// CFC twin of T_SafeEStop_Tests: the same tests drawn as CFC diagrams, the way a TwinSAFE project is authored.
    FUNCTION_BLOCK T_SafeEStop_Tests_CFC EXTENDS T_SafeCfcTestSuite
    VAR
    // Test_OutputsOffWhenStopped
    group_1 : T_SafeGroup;
    fb_1 : T_SafeEStop(group := group_1);
    // Test_StartupRequiresRestartSequence
    group_2 : T_SafeGroup;
    fb_2 : T_SafeEStop(group := group_2);
    // Test_EStopRequestSwitchesOutputsOffAndBlocksRestart
    group_3 : T_SafeGroup;
    fb_3 : T_SafeEStop(group := group_3);
    // Test_MakeContactInputRequestsSafeStateOnOne
    group_4 : T_SafeGroup;
    fb_4 : T_SafeEStop(group := group_4) := (Parameters := (EStopIn1MakeContact := TRUE));
    // Test_EdmErrorAtRestartAndAcknowledge
    group_5 : T_SafeGroup;
    fb_5 : T_SafeEStop(group := group_5);
    // Test_RestartHeldBeforeEStopGivesEdmError
    group_6 : T_SafeGroup;
    fb_6 : T_SafeEStop(group := group_6);
    // Test_DelayedOutput
    group_7 : T_SafeGroup;
    fb_7 : T_SafeEStop(group := group_7) := (Parameters := (DelayTime := T#150MS));
    tR1_7 : TON;
    tR2_7 : TON;
    tPress_7 : TON;
    t1_7 : TON;
    trigPress_7 : R_TRIG;
    trig1_7 : R_TRIG;
    // Test_DiscrepancyErrorNeedsSafeInputsBeforeAck
    group_8 : T_SafeGroup;
    fb_8 : T_SafeEStop(group := group_8) := (Parameters := (DiscrepancyTime1 := T#100MS));
    tR1_8 : TON;
    tR2_8 : TON;
    tPress_8 : TON;
    t1_8 : TON;
    trig1_8 : R_TRIG;
END_VAR

Test_OutputsOffWhenStopped();
Test_StartupRequiresRestartSequence();
Test_EStopRequestSwitchesOutputsOffAndBlocksRestart();
Test_MakeContactInputRequestsSafeStateOnOne();
Test_EdmErrorAtRestartAndAcknowledge();
Test_RestartHeldBeforeEStopGivesEdmError();
Test_DelayedOutput();
Test_DiscrepancyErrorNeedsSafeInputsBeforeAck();

METHOD PRIVATE Test_OutputsOffWhenStopped
// note: this text did not pass the execution check against the stored diagram
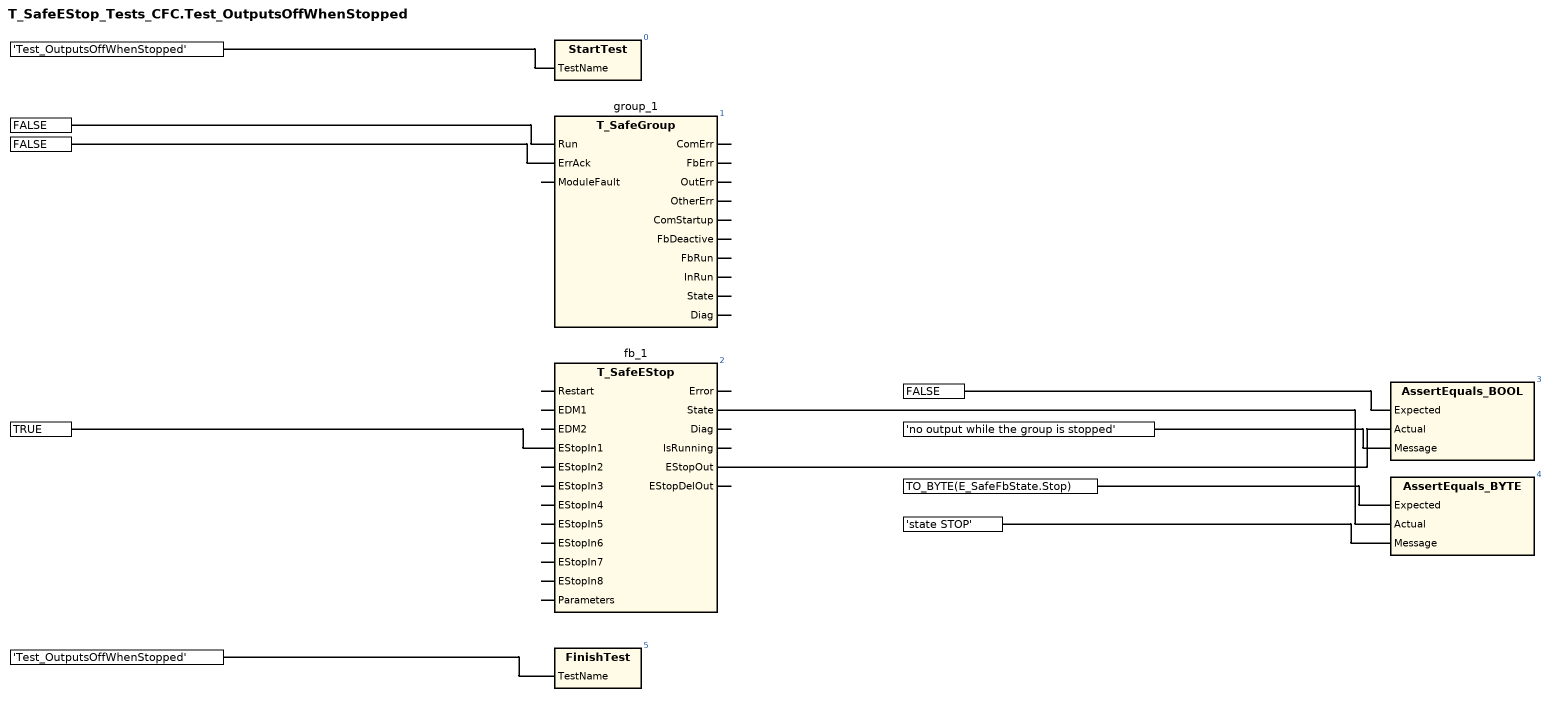
StartTest(TestName := 'Test_OutputsOffWhenStopped');
group_1(Run := FALSE, ErrAck := FALSE); // T_SafeGroup
fb_1(EStopIn1 := TRUE); // T_SafeEStop
AssertEquals_BOOL(Expected := FALSE, Actual := fb_1.EStopOut, Message := 'no output while the group is stopped');
AssertEquals_BYTE(Expected := TO_BYTE(E_SafeFbState.Stop), Actual := fb_1.State, Message := 'state STOP');
FinishTest(TestName := 'Test_OutputsOffWhenStopped');
END_METHOD

METHOD PRIVATE Test_StartupRequiresRestartSequence
// note: this text did not pass the execution check against the stored diagram
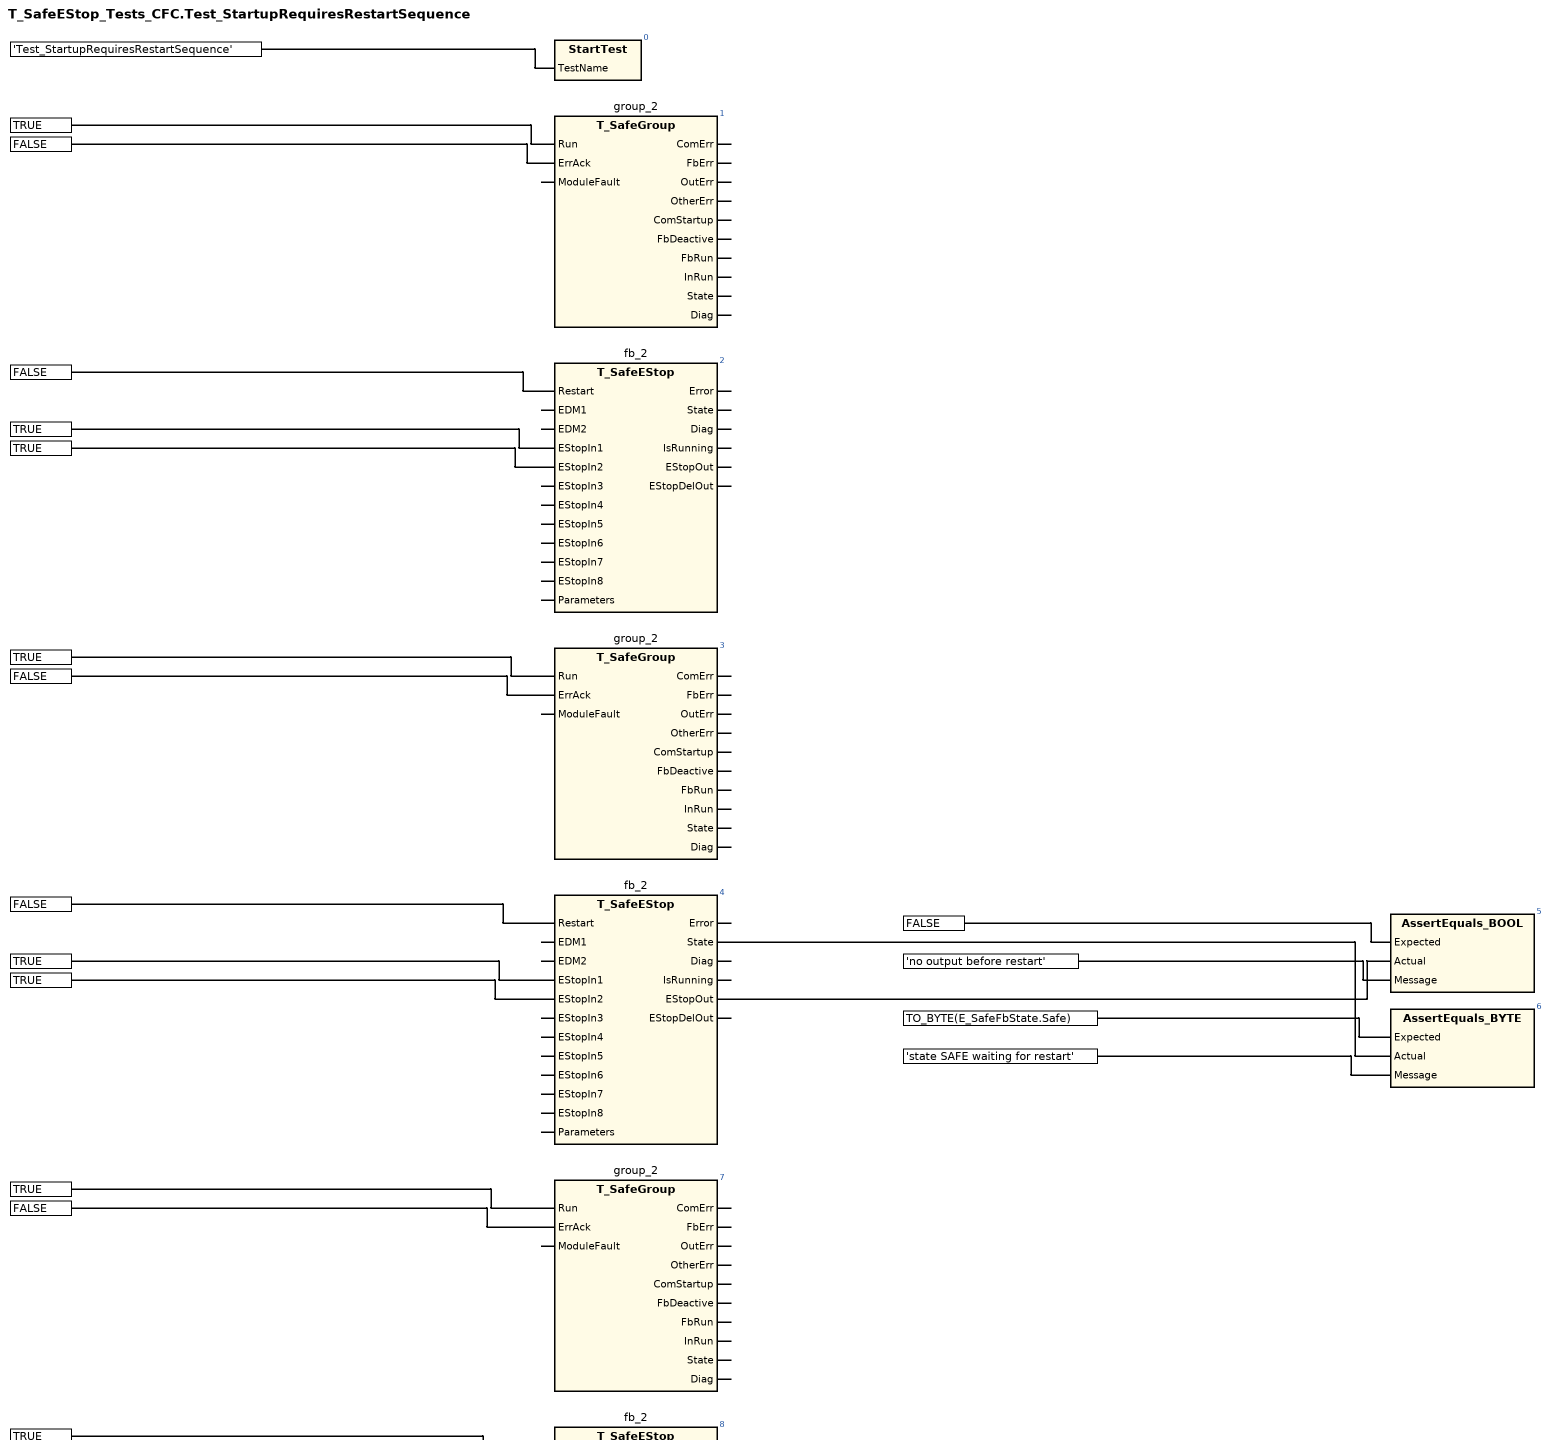
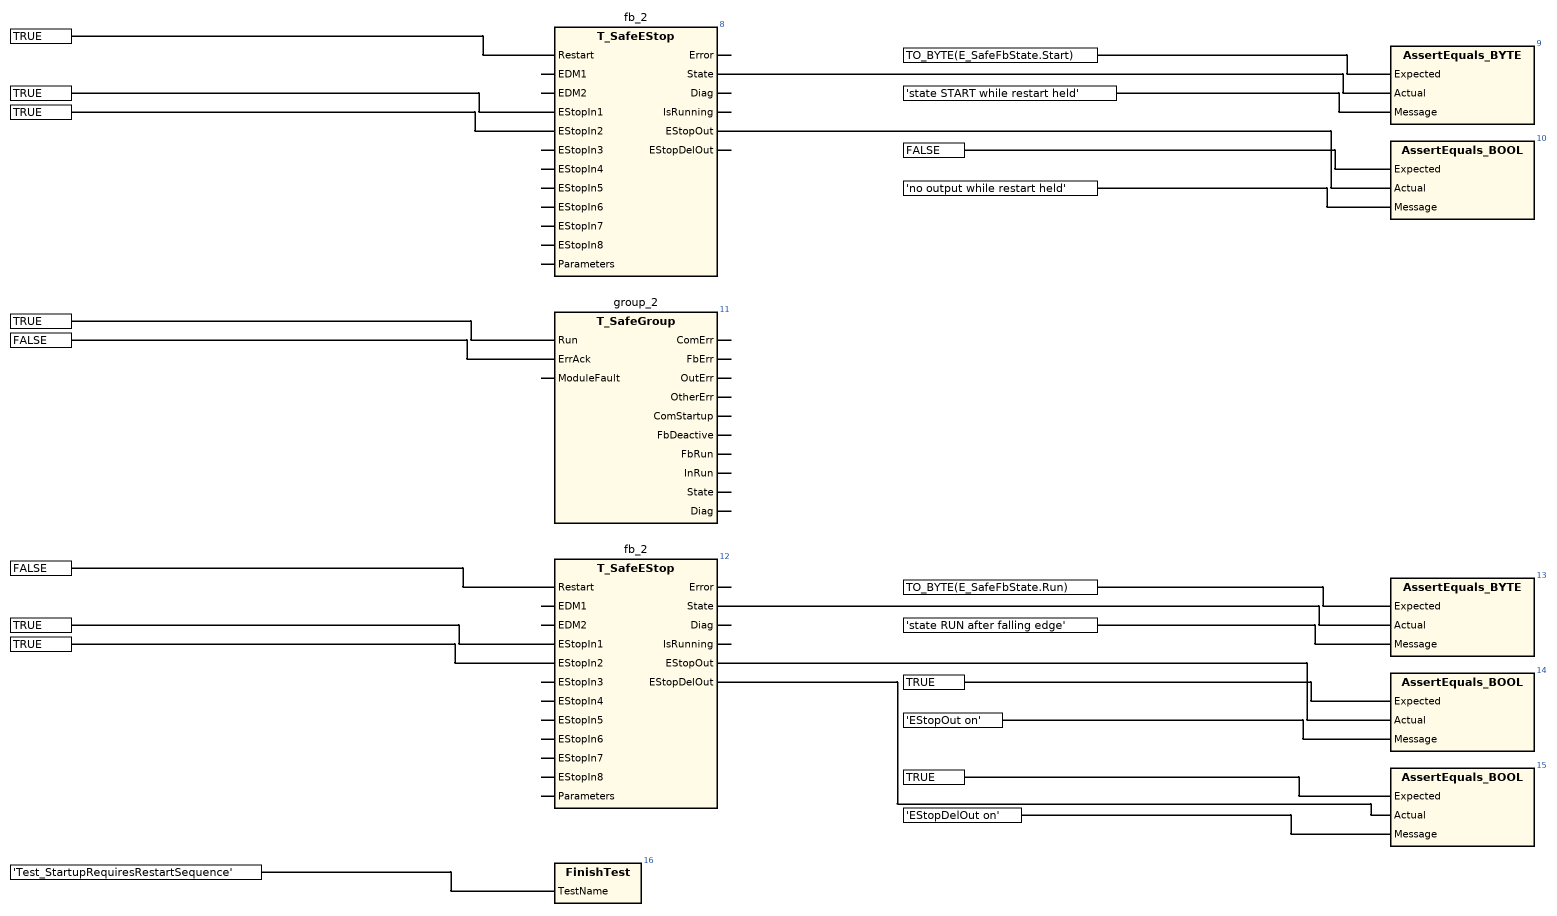
StartTest(TestName := 'Test_StartupRequiresRestartSequence');
group_2(Run := TRUE, ErrAck := FALSE); // T_SafeGroup
fb_2(Restart := FALSE, EStopIn1 := TRUE, EStopIn2 := TRUE); // T_SafeEStop
group_2(Run := TRUE, ErrAck := FALSE); // T_SafeGroup
fb_2(Restart := FALSE, EStopIn1 := TRUE, EStopIn2 := TRUE); // T_SafeEStop
AssertEquals_BOOL(Expected := FALSE, Actual := fb_2.EStopOut, Message := 'no output before restart');
AssertEquals_BYTE(Expected := TO_BYTE(E_SafeFbState.Safe), Actual := fb_2.State, Message := 'state SAFE waiting for restart');
group_2(Run := TRUE, ErrAck := FALSE); // T_SafeGroup
fb_2(Restart := TRUE, EStopIn1 := TRUE, EStopIn2 := TRUE); // T_SafeEStop
AssertEquals_BYTE(Expected := TO_BYTE(E_SafeFbState.Start), Actual := fb_2.State, Message := 'state START while restart held');
AssertEquals_BOOL(Expected := FALSE, Actual := fb_2.EStopOut, Message := 'no output while restart held');
group_2(Run := TRUE, ErrAck := FALSE); // T_SafeGroup
fb_2(Restart := FALSE, EStopIn1 := TRUE, EStopIn2 := TRUE); // T_SafeEStop
AssertEquals_BYTE(Expected := TO_BYTE(E_SafeFbState.Run), Actual := fb_2.State, Message := 'state RUN after falling edge');
AssertEquals_BOOL(Expected := TRUE, Actual := fb_2.EStopOut, Message := 'EStopOut on');
AssertEquals_BOOL(Expected := TRUE, Actual := fb_2.EStopDelOut, Message := 'EStopDelOut on');
FinishTest(TestName := 'Test_StartupRequiresRestartSequence');
END_METHOD

METHOD PRIVATE Test_EStopRequestSwitchesOutputsOffAndBlocksRestart
// note: this text did not pass the execution check against the stored diagram
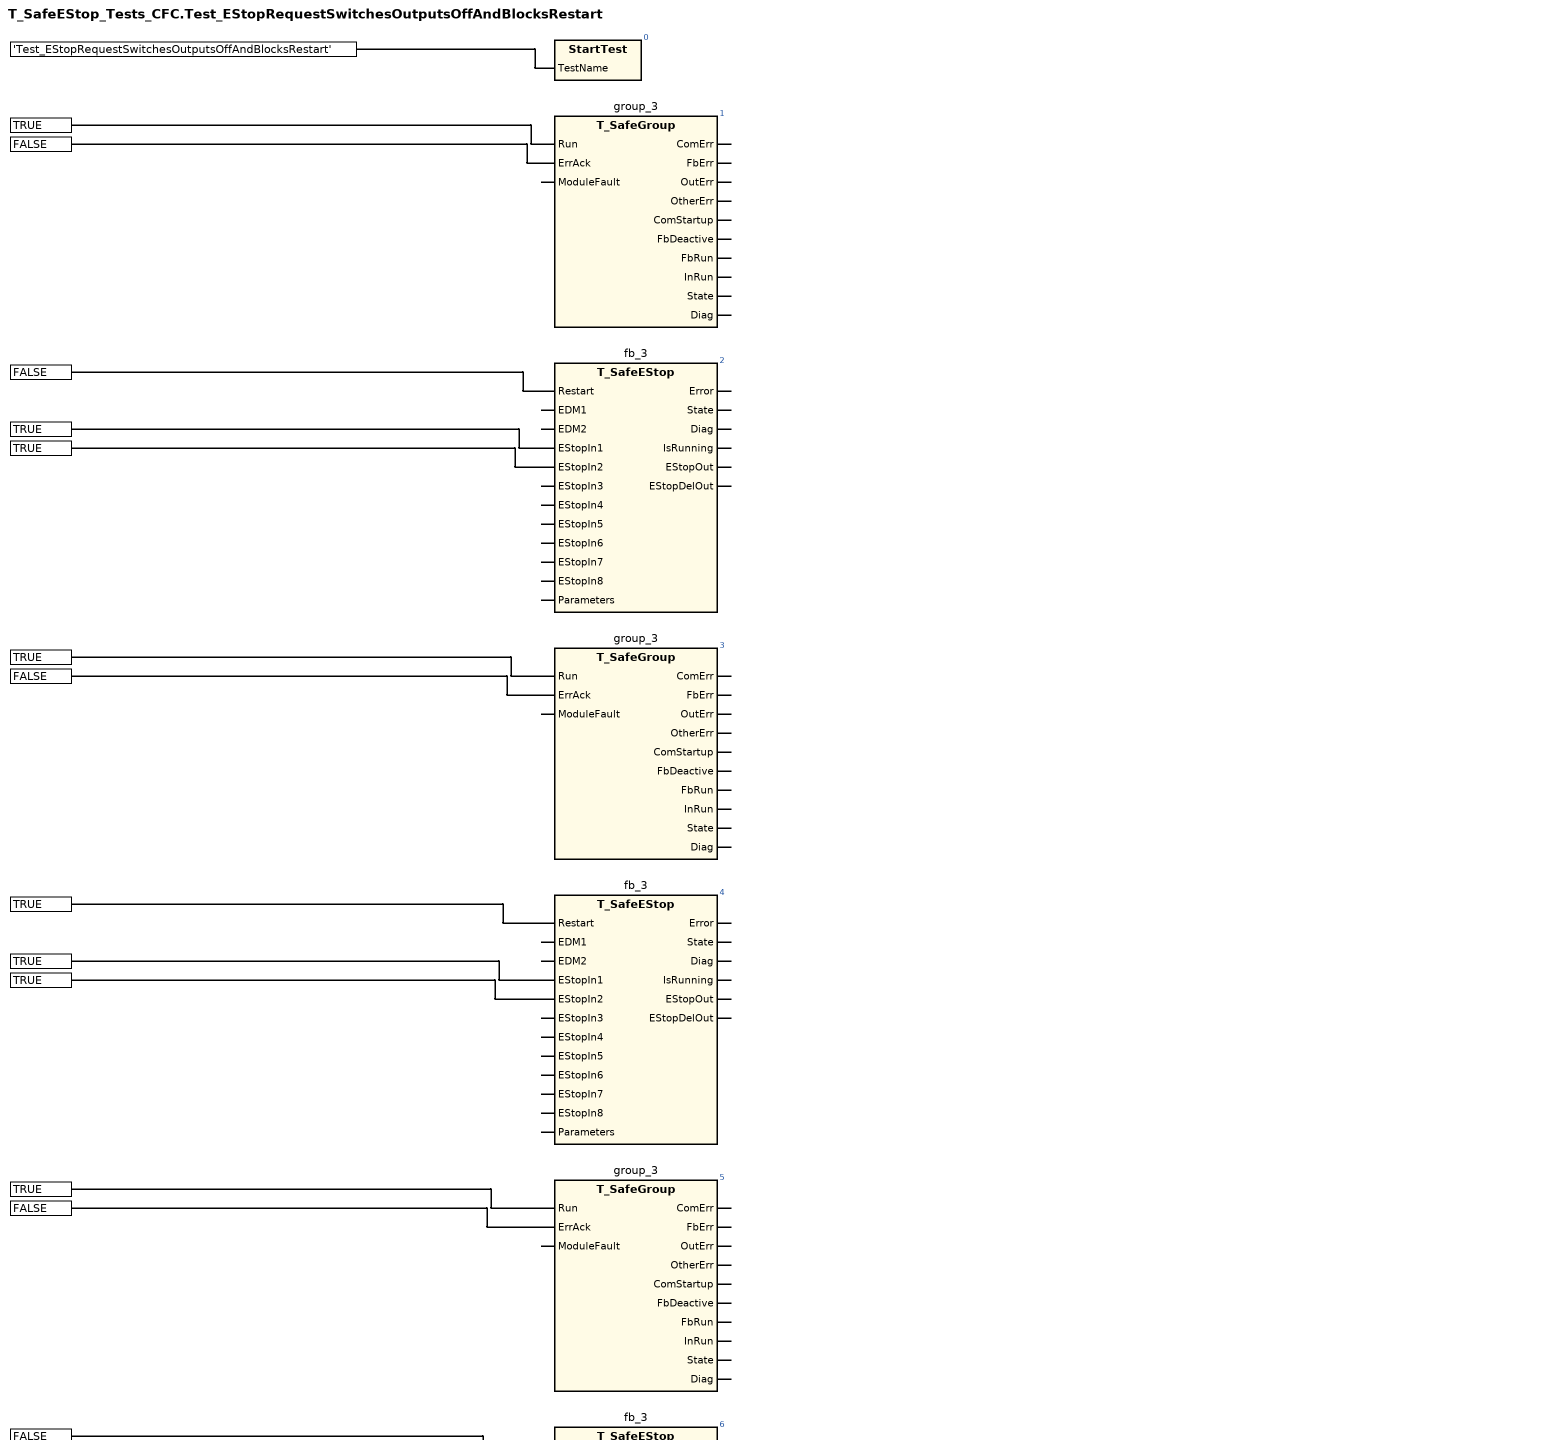
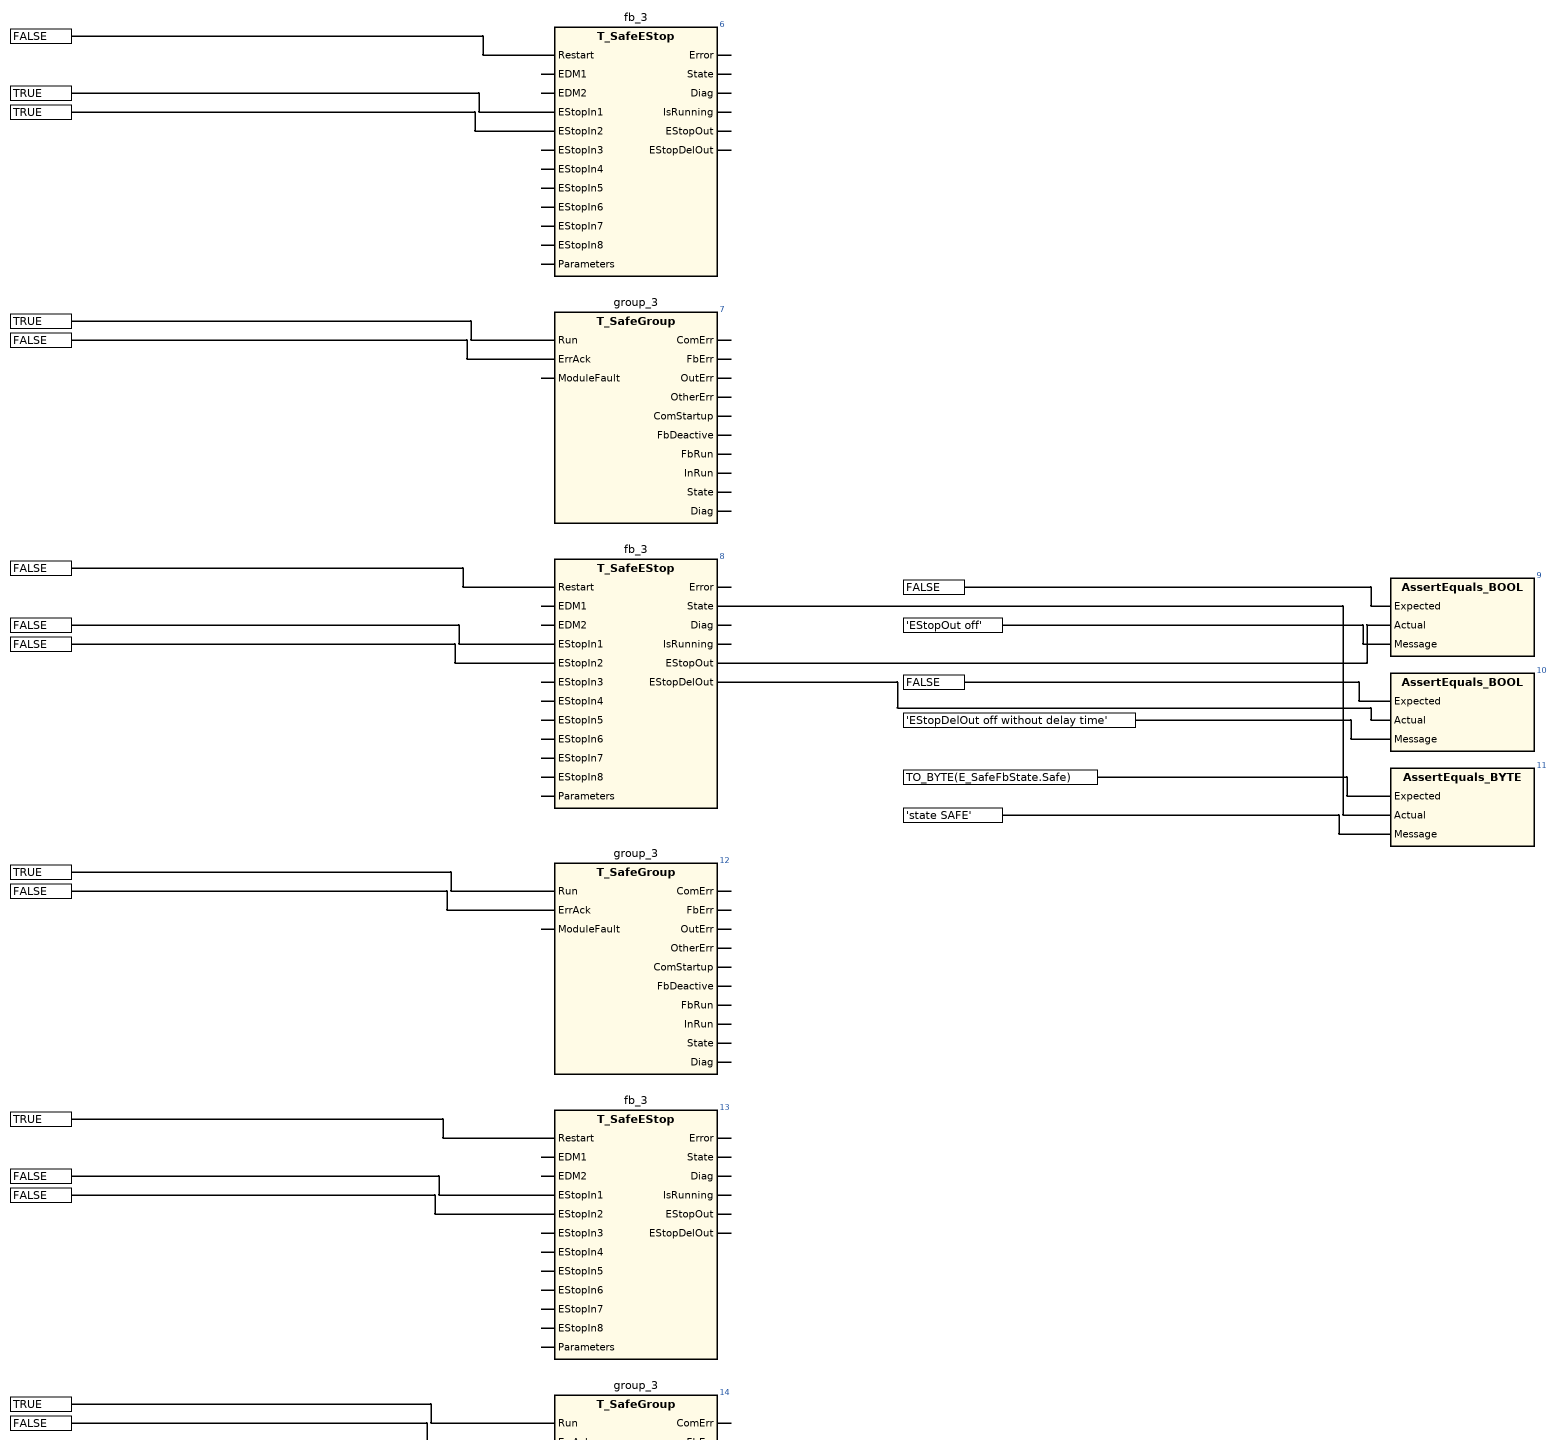
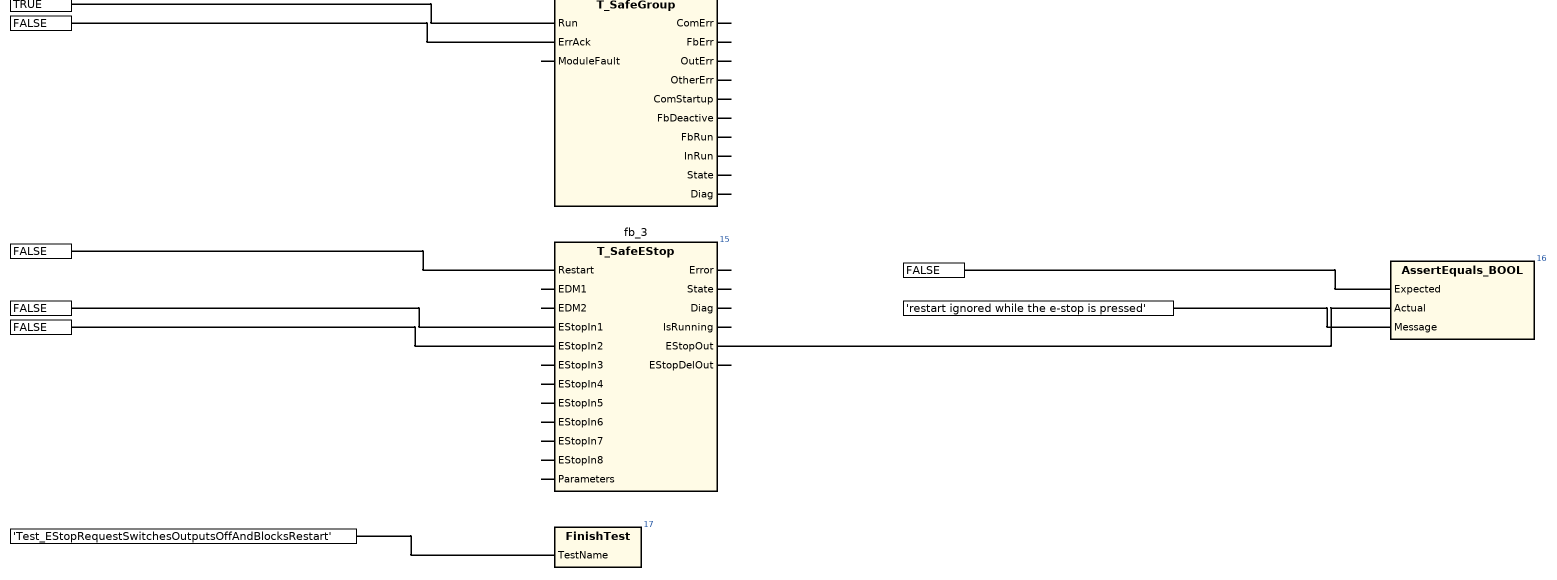
StartTest(TestName := 'Test_EStopRequestSwitchesOutputsOffAndBlocksRestart');
group_3(Run := TRUE, ErrAck := FALSE); // T_SafeGroup
fb_3(Restart := FALSE, EStopIn1 := TRUE, EStopIn2 := TRUE); // T_SafeEStop
group_3(Run := TRUE, ErrAck := FALSE); // T_SafeGroup
fb_3(Restart := TRUE, EStopIn1 := TRUE, EStopIn2 := TRUE); // T_SafeEStop
group_3(Run := TRUE, ErrAck := FALSE); // T_SafeGroup
fb_3(Restart := FALSE, EStopIn1 := TRUE, EStopIn2 := TRUE); // T_SafeEStop
group_3(Run := TRUE, ErrAck := FALSE); // T_SafeGroup
fb_3(Restart := FALSE, EStopIn1 := FALSE, EStopIn2 := FALSE); // T_SafeEStop
AssertEquals_BOOL(Expected := FALSE, Actual := fb_3.EStopOut, Message := 'EStopOut off');
AssertEquals_BOOL(Expected := FALSE, Actual := fb_3.EStopDelOut, Message := 'EStopDelOut off without delay time');
AssertEquals_BYTE(Expected := TO_BYTE(E_SafeFbState.Safe), Actual := fb_3.State, Message := 'state SAFE');
group_3(Run := TRUE, ErrAck := FALSE); // T_SafeGroup
fb_3(Restart := TRUE, EStopIn1 := FALSE, EStopIn2 := FALSE); // T_SafeEStop
group_3(Run := TRUE, ErrAck := FALSE); // T_SafeGroup
fb_3(Restart := FALSE, EStopIn1 := FALSE, EStopIn2 := FALSE); // T_SafeEStop
AssertEquals_BOOL(Expected := FALSE, Actual := fb_3.EStopOut, Message := 'restart ignored while the e-stop is pressed');
FinishTest(TestName := 'Test_EStopRequestSwitchesOutputsOffAndBlocksRestart');
END_METHOD

METHOD PRIVATE Test_MakeContactInputRequestsSafeStateOnOne
// note: this text did not pass the execution check against the stored diagram
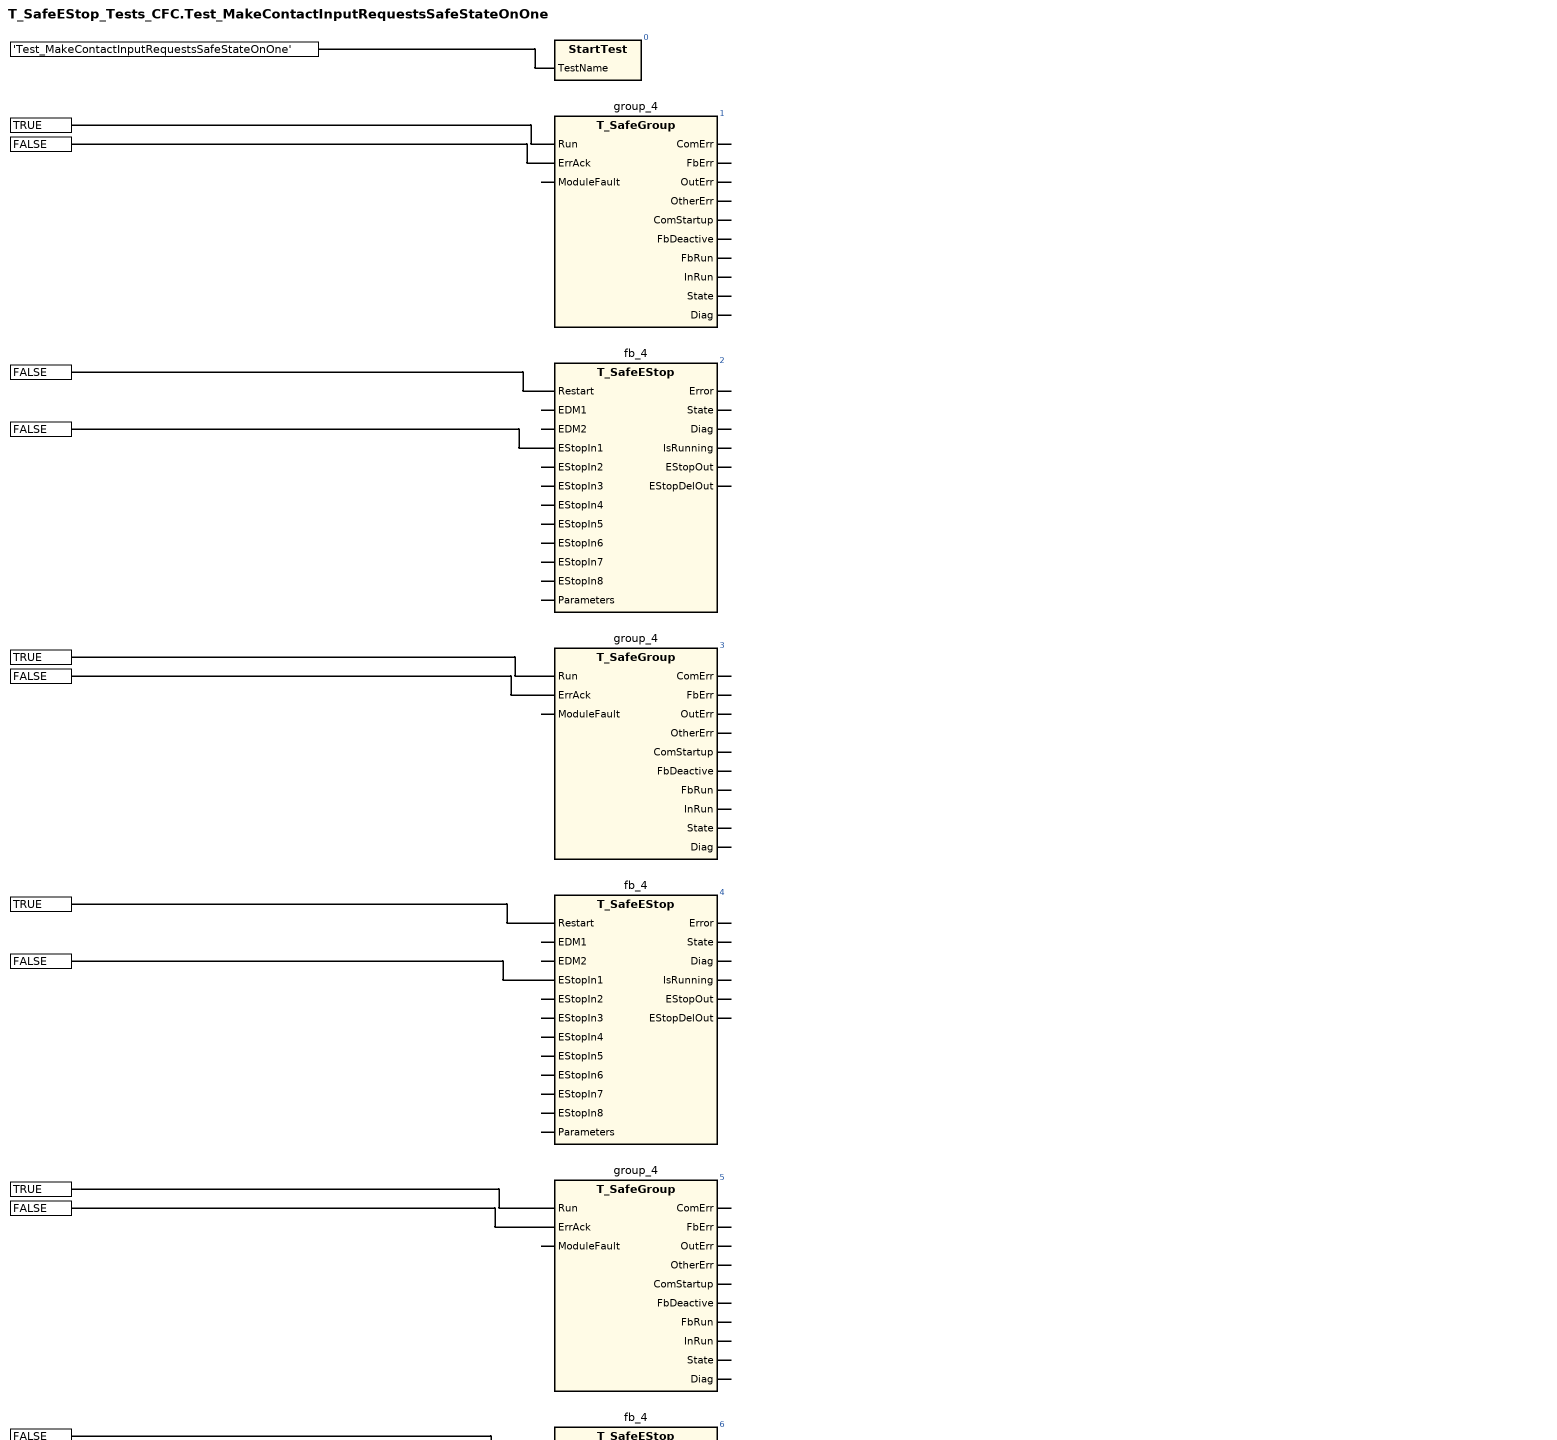
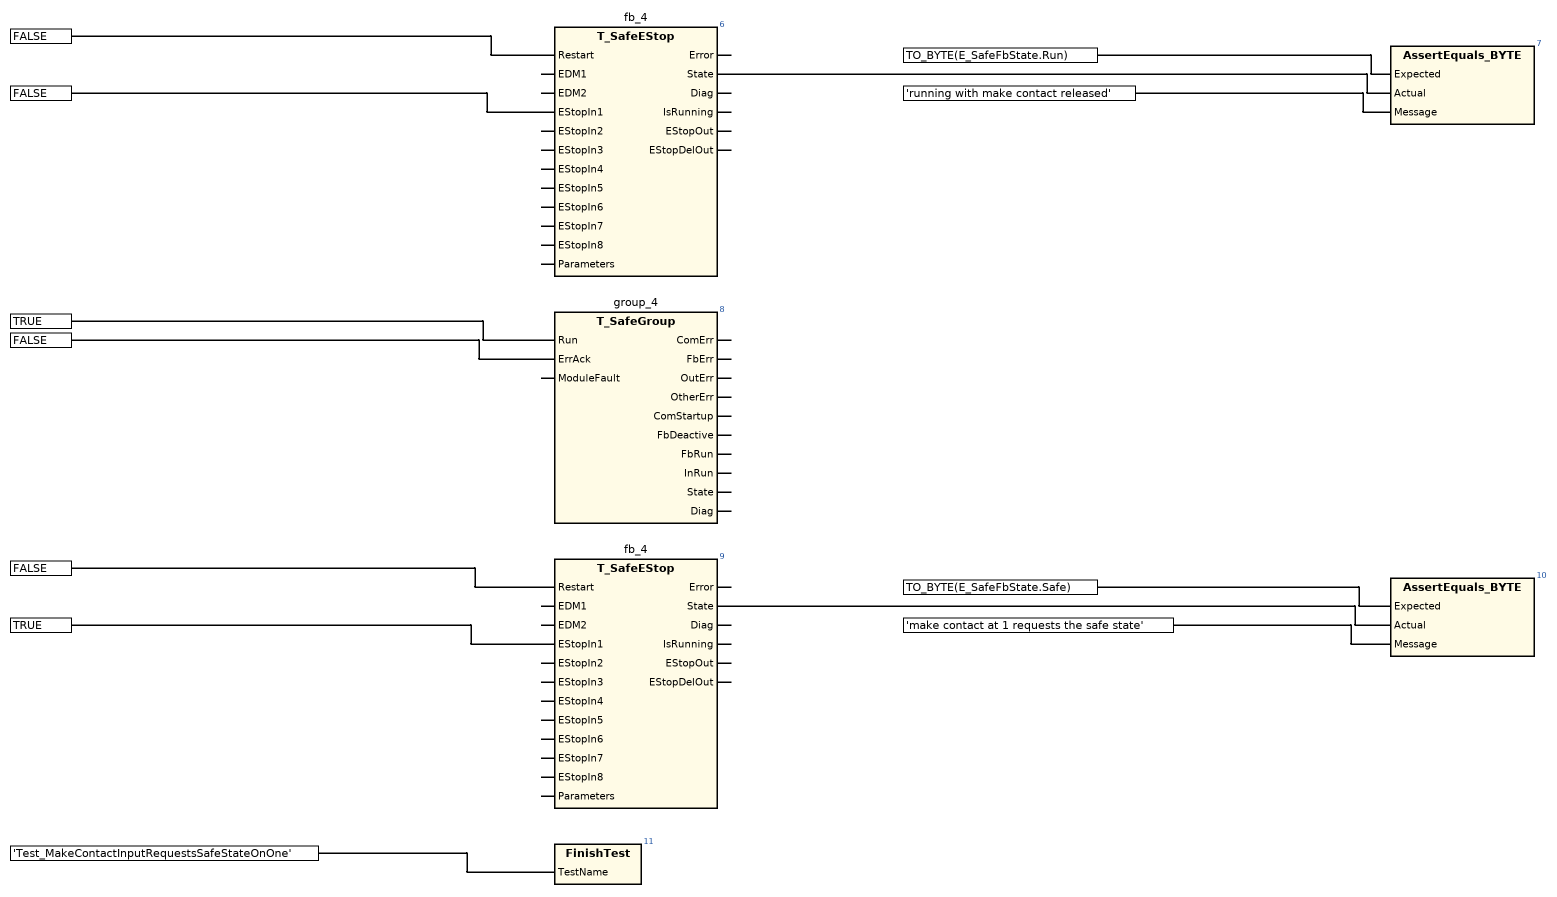
StartTest(TestName := 'Test_MakeContactInputRequestsSafeStateOnOne');
group_4(Run := TRUE, ErrAck := FALSE); // T_SafeGroup
fb_4(Restart := FALSE, EStopIn1 := FALSE); // T_SafeEStop
group_4(Run := TRUE, ErrAck := FALSE); // T_SafeGroup
fb_4(Restart := TRUE, EStopIn1 := FALSE); // T_SafeEStop
group_4(Run := TRUE, ErrAck := FALSE); // T_SafeGroup
fb_4(Restart := FALSE, EStopIn1 := FALSE); // T_SafeEStop
AssertEquals_BYTE(Expected := TO_BYTE(E_SafeFbState.Run), Actual := fb_4.State, Message := 'running with make contact released');
group_4(Run := TRUE, ErrAck := FALSE); // T_SafeGroup
fb_4(Restart := FALSE, EStopIn1 := TRUE); // T_SafeEStop
AssertEquals_BYTE(Expected := TO_BYTE(E_SafeFbState.Safe), Actual := fb_4.State, Message := 'make contact at 1 requests the safe state');
FinishTest(TestName := 'Test_MakeContactInputRequestsSafeStateOnOne');
END_METHOD

METHOD PRIVATE Test_EdmErrorAtRestartAndAcknowledge
// note: this text did not pass the execution check against the stored diagram
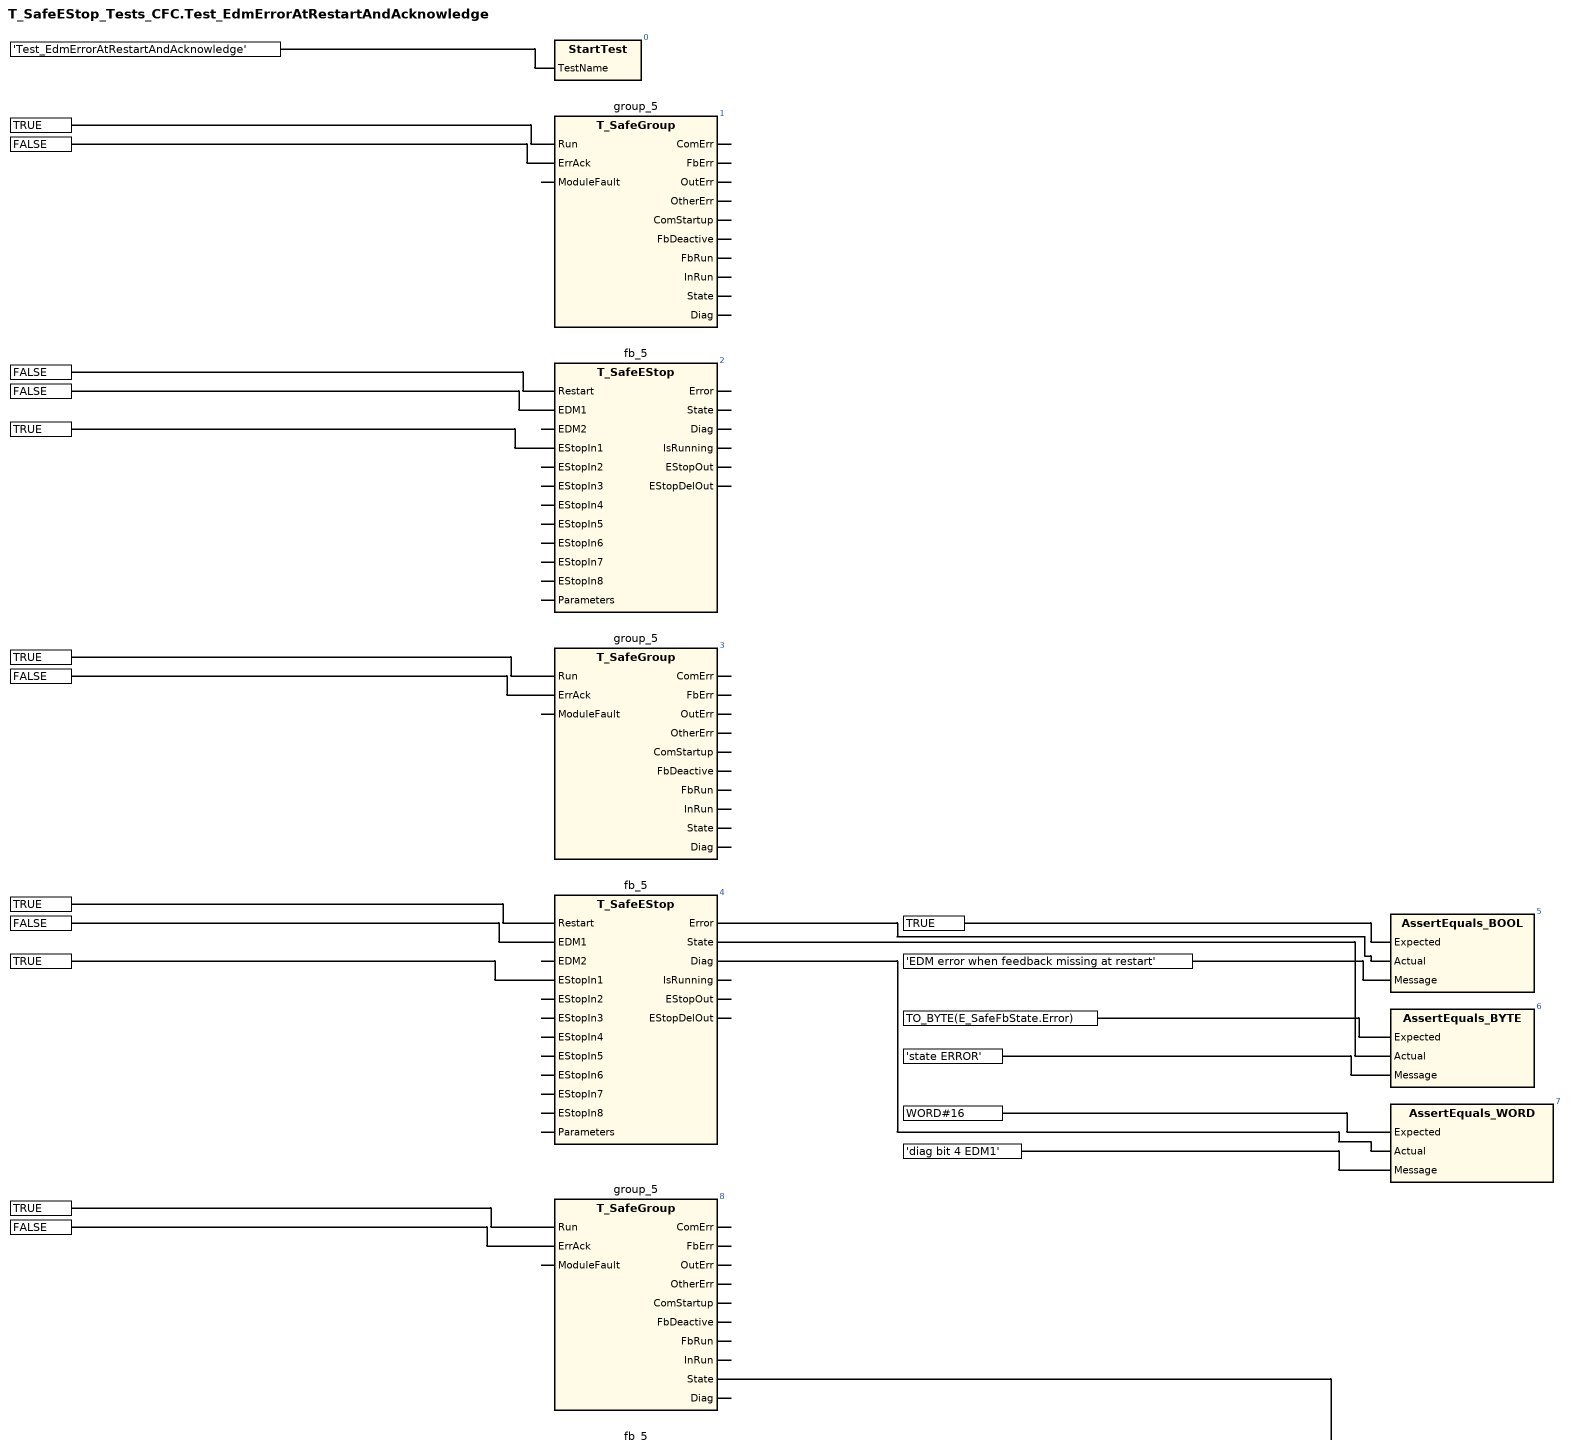
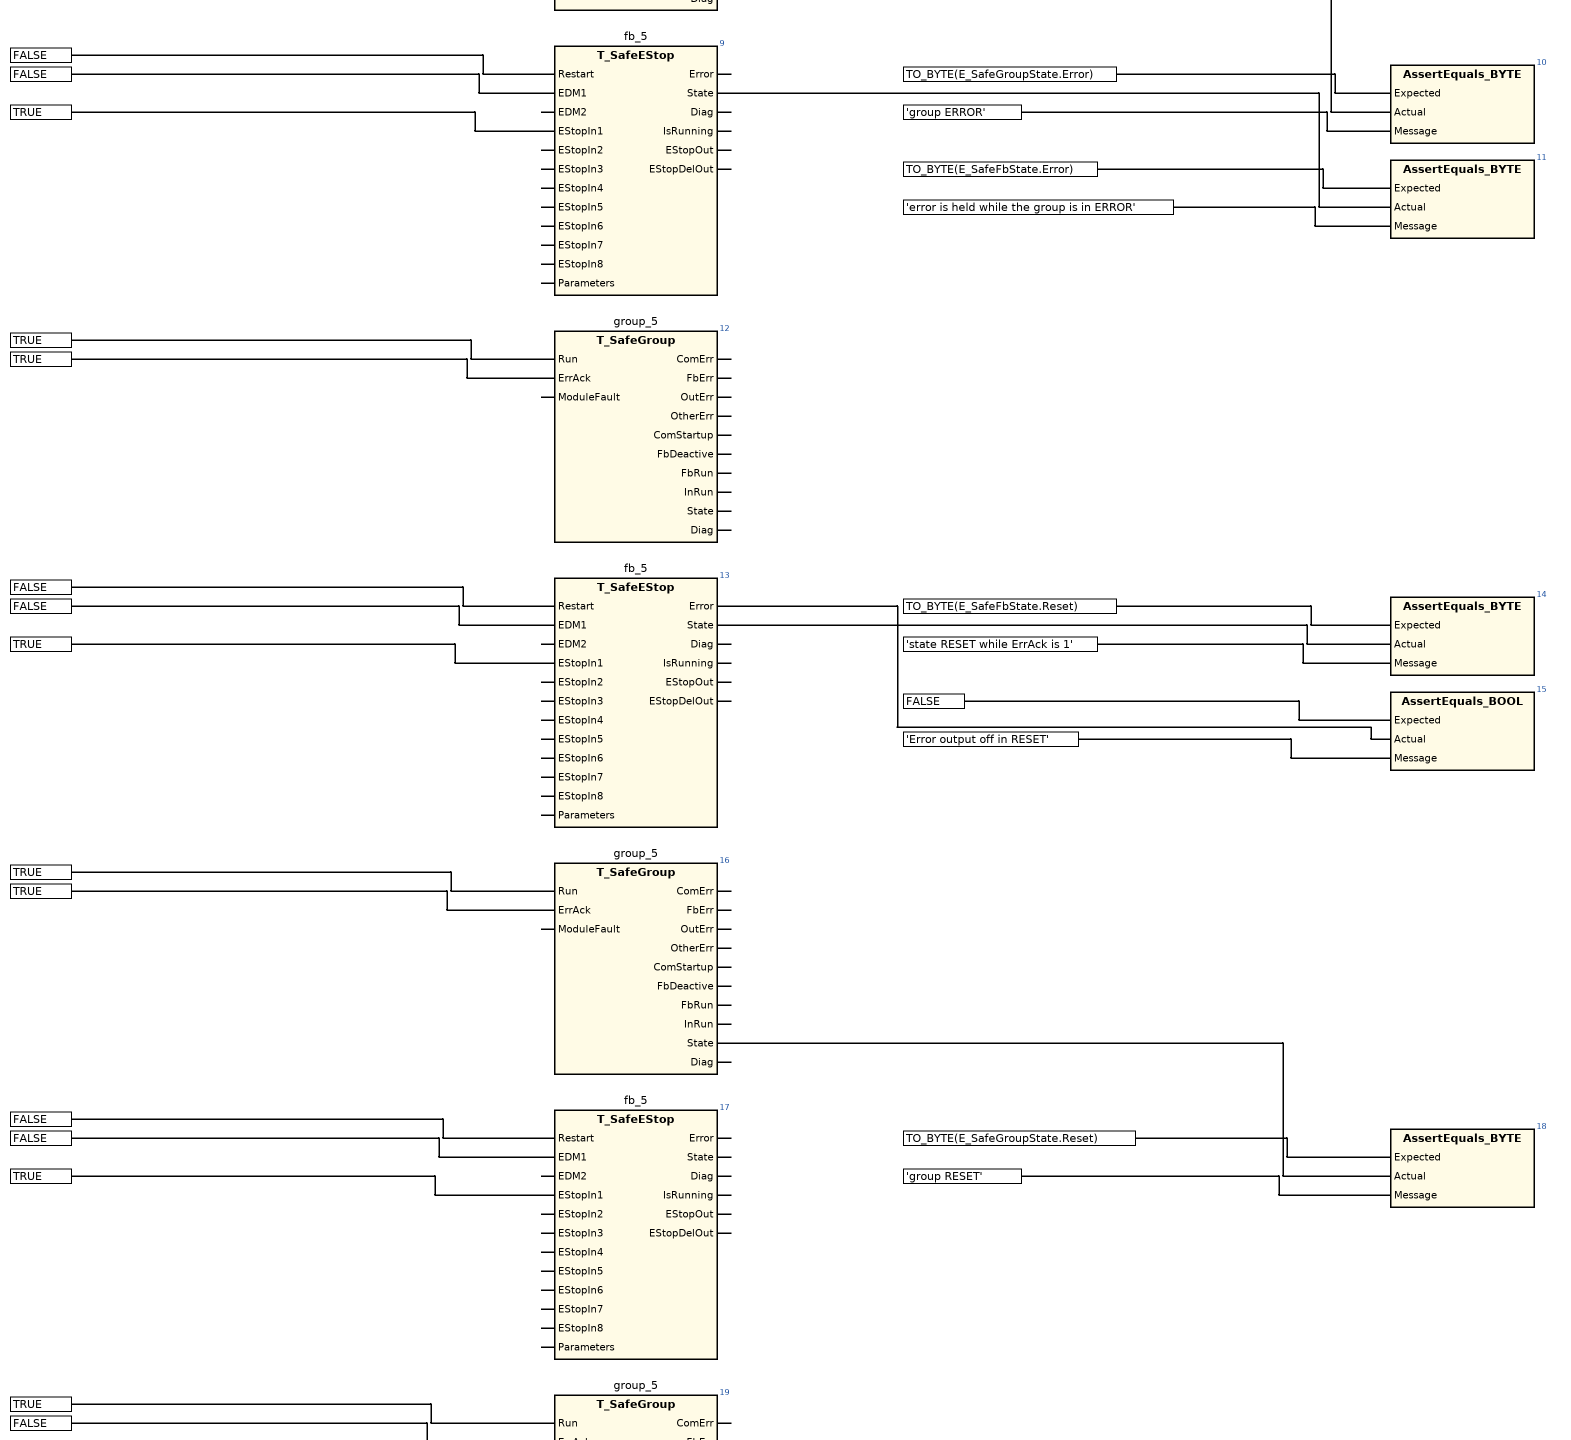
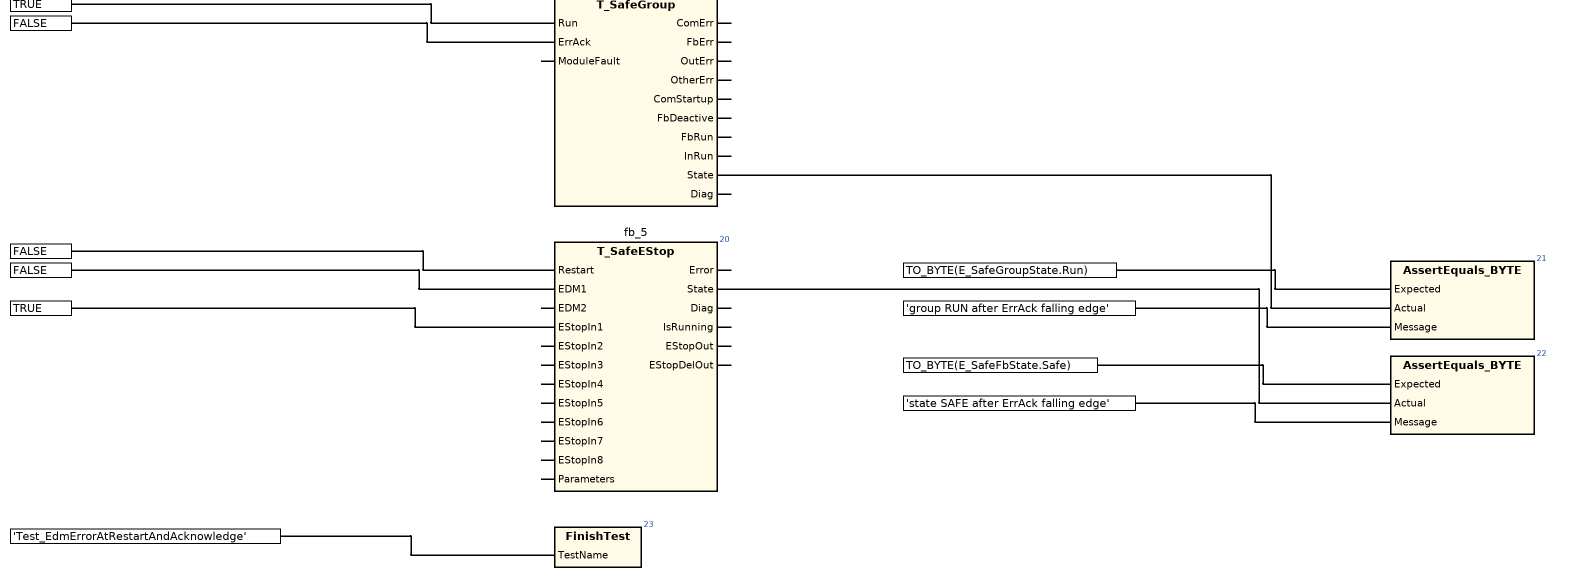
StartTest(TestName := 'Test_EdmErrorAtRestartAndAcknowledge');
group_5(Run := TRUE, ErrAck := FALSE); // T_SafeGroup
fb_5(Restart := FALSE, EDM1 := FALSE, EStopIn1 := TRUE); // T_SafeEStop
group_5(Run := TRUE, ErrAck := FALSE); // T_SafeGroup
fb_5(Restart := TRUE, EDM1 := FALSE, EStopIn1 := TRUE); // T_SafeEStop
AssertEquals_BOOL(Expected := TRUE, Actual := fb_5.Error, Message := 'EDM error when feedback missing at restart');
AssertEquals_BYTE(Expected := TO_BYTE(E_SafeFbState.Error), Actual := fb_5.State, Message := 'state ERROR');
AssertEquals_WORD(Expected := WORD#16, Actual := fb_5.Diag, Message := 'diag bit 4 EDM1');
group_5(Run := TRUE, ErrAck := FALSE); // T_SafeGroup
fb_5(Restart := FALSE, EDM1 := FALSE, EStopIn1 := TRUE); // T_SafeEStop
AssertEquals_BYTE(Expected := TO_BYTE(E_SafeGroupState.Error), Actual := group_5.State, Message := 'group ERROR');
AssertEquals_BYTE(Expected := TO_BYTE(E_SafeFbState.Error), Actual := fb_5.State, Message := 'error is held while the group is in ERROR');
group_5(Run := TRUE, ErrAck := TRUE); // T_SafeGroup
fb_5(Restart := FALSE, EDM1 := FALSE, EStopIn1 := TRUE); // T_SafeEStop
AssertEquals_BYTE(Expected := TO_BYTE(E_SafeFbState.Reset), Actual := fb_5.State, Message := 'state RESET while ErrAck is 1');
AssertEquals_BOOL(Expected := FALSE, Actual := fb_5.Error, Message := 'Error output off in RESET');
group_5(Run := TRUE, ErrAck := TRUE); // T_SafeGroup
fb_5(Restart := FALSE, EDM1 := FALSE, EStopIn1 := TRUE); // T_SafeEStop
AssertEquals_BYTE(Expected := TO_BYTE(E_SafeGroupState.Reset), Actual := group_5.State, Message := 'group RESET');
group_5(Run := TRUE, ErrAck := FALSE); // T_SafeGroup
fb_5(Restart := FALSE, EDM1 := FALSE, EStopIn1 := TRUE); // T_SafeEStop
AssertEquals_BYTE(Expected := TO_BYTE(E_SafeGroupState.Run), Actual := group_5.State, Message := 'group RUN after ErrAck falling edge');
AssertEquals_BYTE(Expected := TO_BYTE(E_SafeFbState.Safe), Actual := fb_5.State, Message := 'state SAFE after ErrAck falling edge');
FinishTest(TestName := 'Test_EdmErrorAtRestartAndAcknowledge');
END_METHOD

METHOD PRIVATE Test_RestartHeldBeforeEStopGivesEdmError
// note: this text did not pass the execution check against the stored diagram
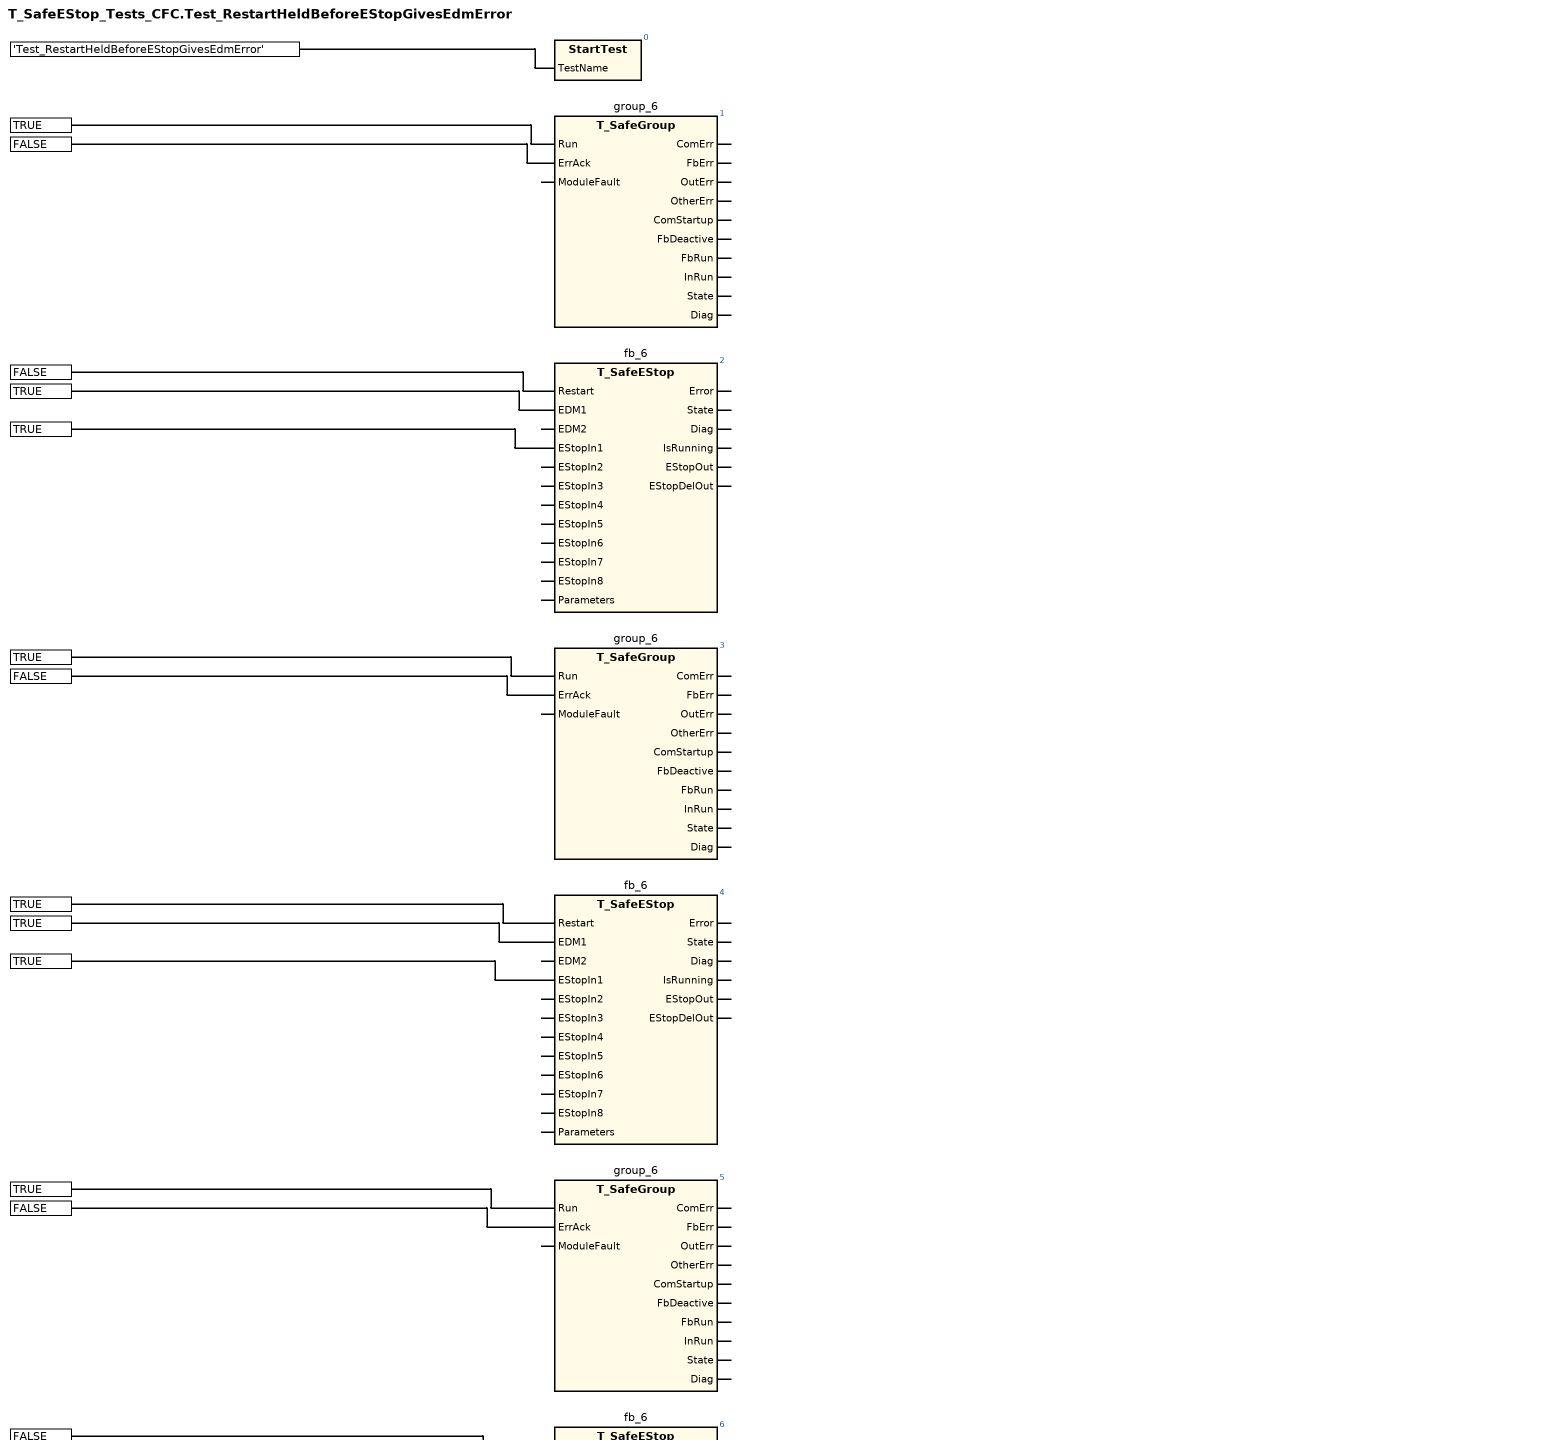
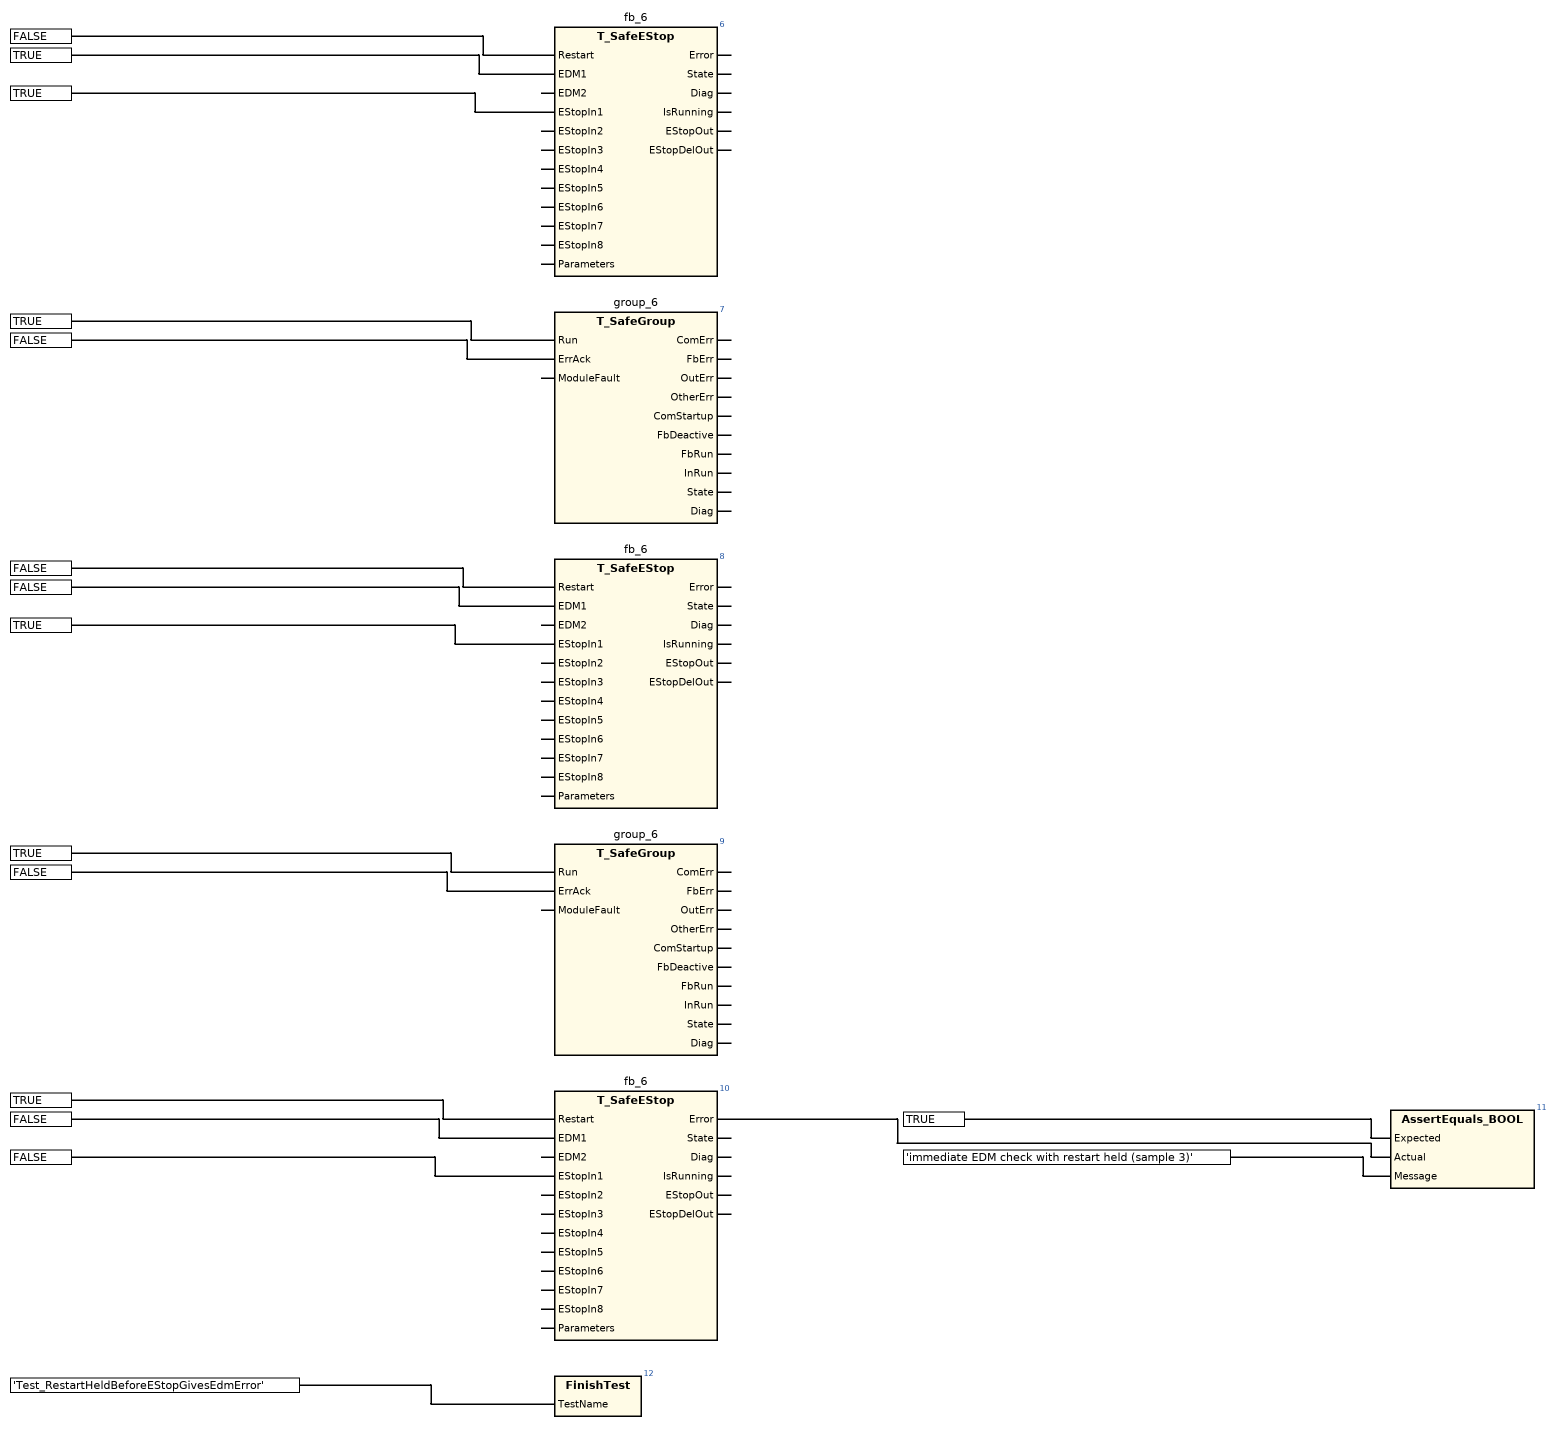
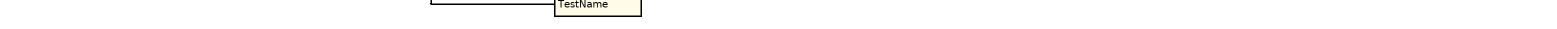
StartTest(TestName := 'Test_RestartHeldBeforeEStopGivesEdmError');
group_6(Run := TRUE, ErrAck := FALSE); // T_SafeGroup
fb_6(Restart := FALSE, EDM1 := TRUE, EStopIn1 := TRUE); // T_SafeEStop
group_6(Run := TRUE, ErrAck := FALSE); // T_SafeGroup
fb_6(Restart := TRUE, EDM1 := TRUE, EStopIn1 := TRUE); // T_SafeEStop
group_6(Run := TRUE, ErrAck := FALSE); // T_SafeGroup
fb_6(Restart := FALSE, EDM1 := TRUE, EStopIn1 := TRUE); // T_SafeEStop
group_6(Run := TRUE, ErrAck := FALSE); // T_SafeGroup
fb_6(Restart := FALSE, EDM1 := FALSE, EStopIn1 := TRUE); // T_SafeEStop
group_6(Run := TRUE, ErrAck := FALSE); // T_SafeGroup
fb_6(Restart := TRUE, EDM1 := FALSE, EStopIn1 := FALSE); // T_SafeEStop
AssertEquals_BOOL(Expected := TRUE, Actual := fb_6.Error, Message := 'immediate EDM check with restart held (sample 3)');
FinishTest(TestName := 'Test_RestartHeldBeforeEStopGivesEdmError');
END_METHOD

METHOD PRIVATE Test_DelayedOutput
// note: this text did not pass the execution check against the stored diagram
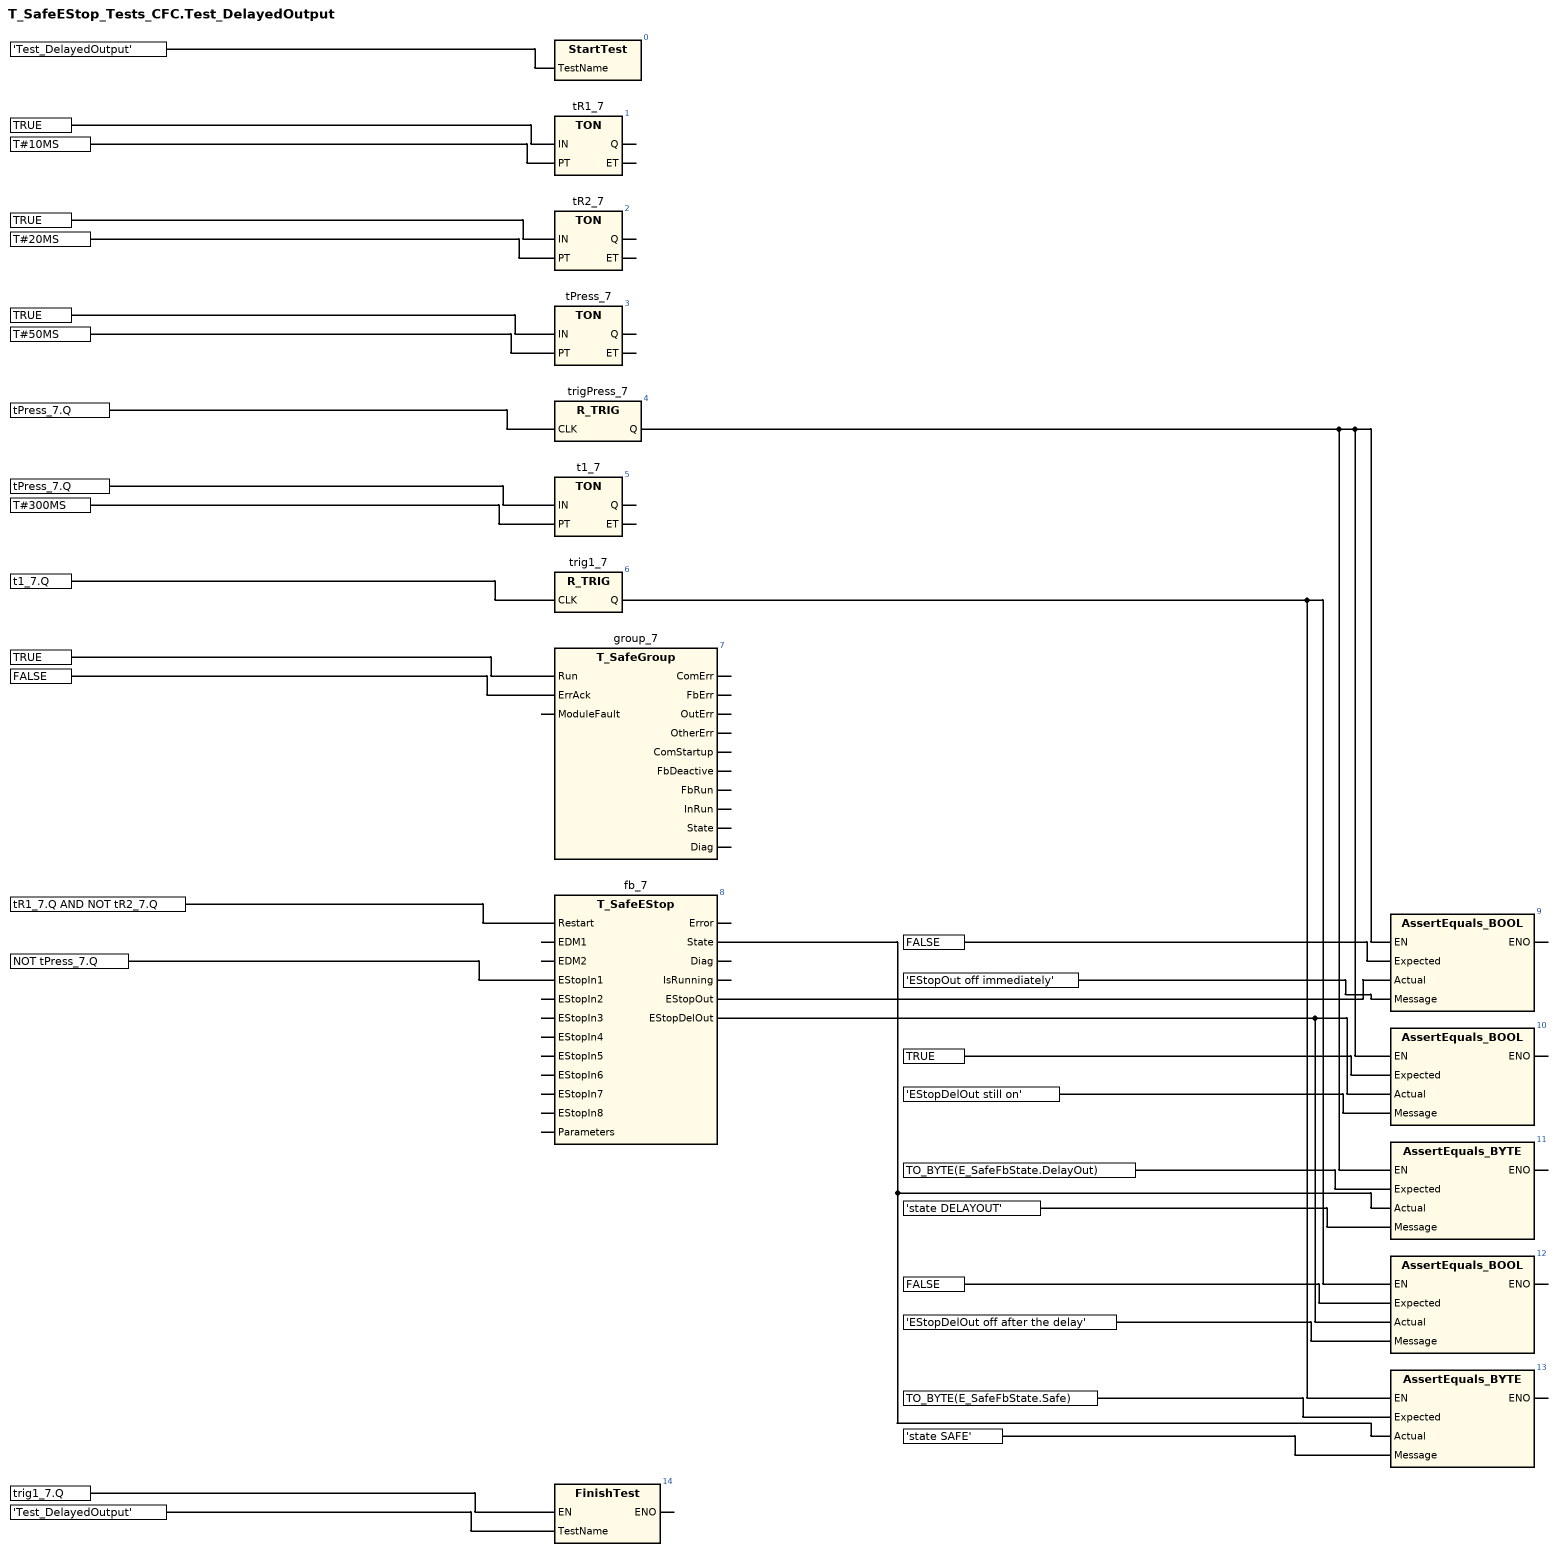
StartTest(TestName := 'Test_DelayedOutput');
tR1_7(IN := TRUE, PT := T#10MS); // TON
tR2_7(IN := TRUE, PT := T#20MS); // TON
tPress_7(IN := TRUE, PT := T#50MS); // TON
trigPress_7(CLK := tPress_7.Q); // R_TRIG
t1_7(IN := tPress_7.Q, PT := T#300MS); // TON
trig1_7(CLK := t1_7.Q); // R_TRIG
group_7(Run := TRUE, ErrAck := FALSE); // T_SafeGroup
fb_7(Restart := tR1_7.Q AND NOT tR2_7.Q, EStopIn1 := NOT tPress_7.Q); // T_SafeEStop
IF trigPress_7.Q THEN AssertEquals_BOOL(Expected := FALSE, Actual := fb_7.EStopOut, Message := 'EStopOut off immediately'); END_IF
IF trigPress_7.Q THEN AssertEquals_BOOL(Expected := TRUE, Actual := fb_7.EStopDelOut, Message := 'EStopDelOut still on'); END_IF
IF trigPress_7.Q THEN AssertEquals_BYTE(Expected := TO_BYTE(E_SafeFbState.DelayOut), Actual := fb_7.State, Message := 'state DELAYOUT'); END_IF
IF trig1_7.Q THEN AssertEquals_BOOL(Expected := FALSE, Actual := fb_7.EStopDelOut, Message := 'EStopDelOut off after the delay'); END_IF
IF trig1_7.Q THEN AssertEquals_BYTE(Expected := TO_BYTE(E_SafeFbState.Safe), Actual := fb_7.State, Message := 'state SAFE'); END_IF
IF trig1_7.Q THEN FinishTest(TestName := 'Test_DelayedOutput'); END_IF
END_METHOD

METHOD PRIVATE Test_DiscrepancyErrorNeedsSafeInputsBeforeAck
// note: this text did not pass the execution check against the stored diagram
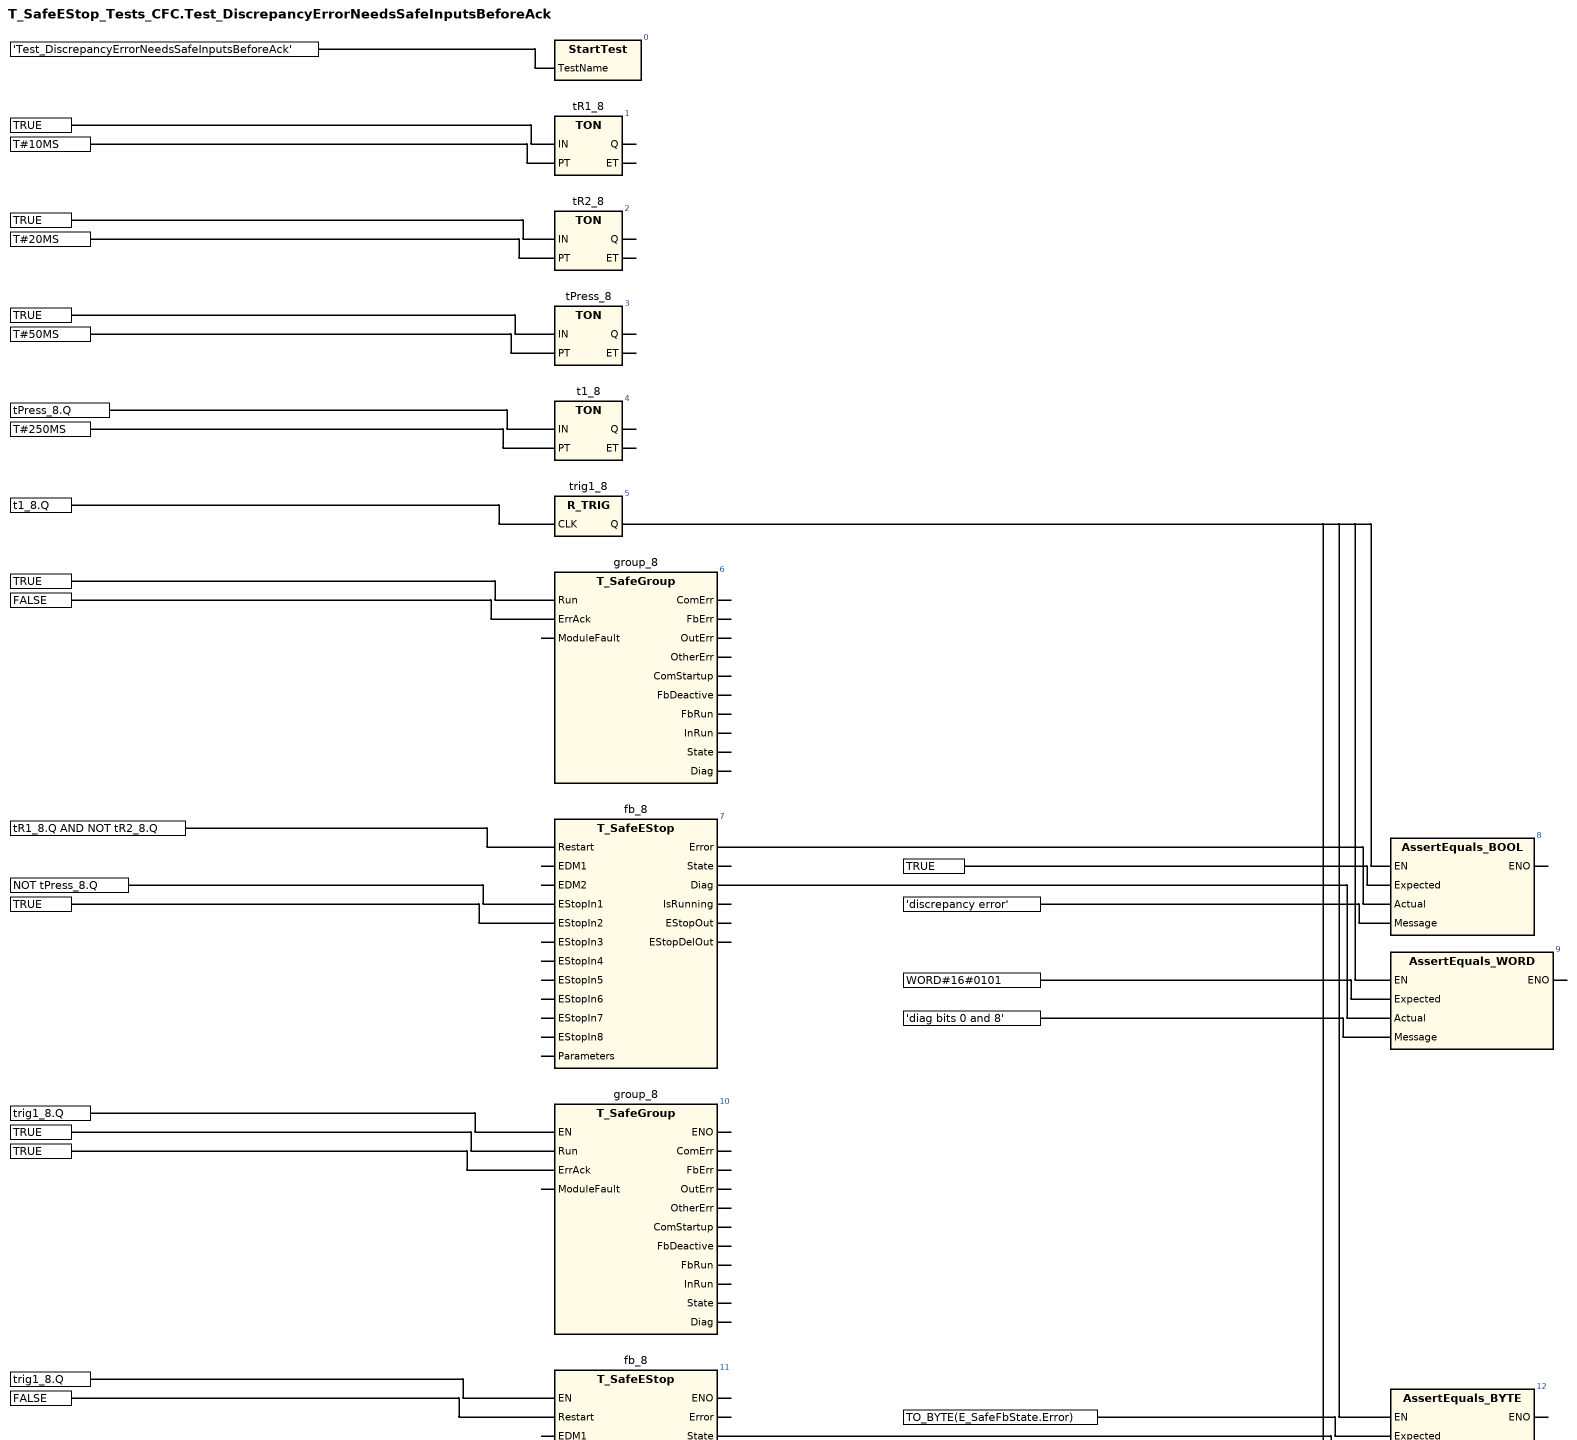
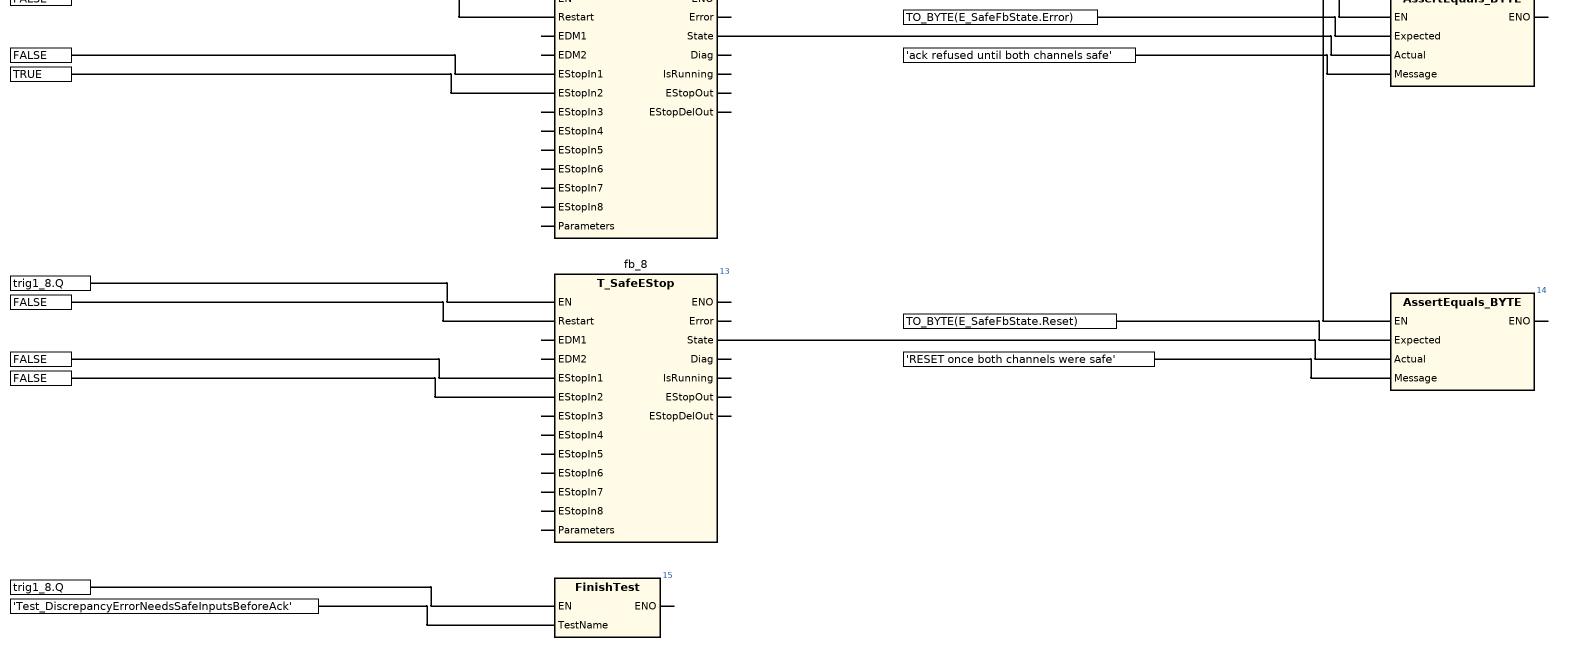
StartTest(TestName := 'Test_DiscrepancyErrorNeedsSafeInputsBeforeAck');
tR1_8(IN := TRUE, PT := T#10MS); // TON
tR2_8(IN := TRUE, PT := T#20MS); // TON
tPress_8(IN := TRUE, PT := T#50MS); // TON
t1_8(IN := tPress_8.Q, PT := T#250MS); // TON
trig1_8(CLK := t1_8.Q); // R_TRIG
group_8(Run := TRUE, ErrAck := FALSE); // T_SafeGroup
fb_8(Restart := tR1_8.Q AND NOT tR2_8.Q, EStopIn1 := NOT tPress_8.Q, EStopIn2 := TRUE); // T_SafeEStop
IF trig1_8.Q THEN AssertEquals_BOOL(Expected := TRUE, Actual := fb_8.Error, Message := 'discrepancy error'); END_IF
IF trig1_8.Q THEN AssertEquals_WORD(Expected := WORD#16#0101, Actual := fb_8.Diag, Message := 'diag bits 0 and 8'); END_IF
IF trig1_8.Q THEN
    group_8(Run := TRUE, ErrAck := TRUE); // T_SafeGroup
END_IF
IF trig1_8.Q THEN
    fb_8(Restart := FALSE, EStopIn1 := FALSE, EStopIn2 := TRUE); // T_SafeEStop
END_IF
IF trig1_8.Q THEN AssertEquals_BYTE(Expected := TO_BYTE(E_SafeFbState.Error), Actual := fb_8.State, Message := 'ack refused until both channels safe'); END_IF
IF trig1_8.Q THEN
    fb_8(Restart := FALSE, EStopIn1 := FALSE, EStopIn2 := FALSE); // T_SafeEStop
END_IF
IF trig1_8.Q THEN AssertEquals_BYTE(Expected := TO_BYTE(E_SafeFbState.Reset), Actual := fb_8.State, Message := 'RESET once both channels were safe'); END_IF
IF trig1_8.Q THEN FinishTest(TestName := 'Test_DiscrepancyErrorNeedsSafeInputsBeforeAck'); END_IF
END_METHOD

END_FUNCTION_BLOCK

(* stored: Version 1.1.0.1, ProductVersion 3.1.4026.22
   POU T_SafeEStop_Tests_CFC: Id {b635a8d4-cc9f-50c7-a7cf-809816fd247d}, SpecialFunc None
   Method Test_OutputsOffWhenStopped: Id {6911d1c7-9bc1-5e3c-8f0b-a41c885fe702}
   Method Test_StartupRequiresRestartSequence: Id {60a7f7f7-6b6f-52ef-b577-763e4f21c945}
   Method Test_EStopRequestSwitchesOutputsOffAndBlocksRestart: Id {4abb9636-3416-53e3-9917-720540bee31a}
   Method Test_MakeContactInputRequestsSafeStateOnOne: Id {4c9b63d5-e9f0-5cc4-a9d0-0eb3581ff610}
   Method Test_EdmErrorAtRestartAndAcknowledge: Id {0f387f1b-bdc6-54ff-8844-74959a5c3a71}
   Method Test_RestartHeldBeforeEStopGivesEdmError: Id {87df58b8-c27b-5571-ba38-9a3de28d8d06}
   Method Test_DelayedOutput: Id {1d167897-cc51-54c8-aaf0-74b6b2a8cd9f}
   Method Test_DiscrepancyErrorNeedsSafeInputsBeforeAck: Id {5609898b-41e9-593d-af57-b1a25f7b531d} *)
